FUNCTION_BLOCK "FB5002_SafetyDoorV1"   // FB5002, SCL
{ S7_Optimized_Access := 'TRUE' }
// ============================================================
//  Block: FB5002_SafetyDoorV1
//  ============================================================
//  编号：FB5002
//  原始语言：LAD（规则翻译为 SCL）
//  含义：由 LAD/FBD 网络折叠生成的等效 SCL，导入前请人工复核
   VAR_INPUT
      i_DoorOverRide : Bool;   // 安全门旁路输入请求信号
      i_AutoRunning : Bool;   // 自动运行中
      i_OpenDoorPmt : Bool := TRUE;   // 开门/旁路条件
      EMMode : Bool;   // 紧急停止模式
   END_VAR
   VAR_OUTPUT
      o_DoorOverRideRelayOn : Bool;   // 安全门旁路继电器输出
      o_DoorLockRelayON : Bool;   // 安全门线圈锁定继电器输出
      o_DoorOverRideLight : Bool;   // 安全门旁路指示灯
      o_PromptDoorOverRideStartIng : Bool;   // 开始安全门旁路,等待各流程结束!
      o_PromptDoorOveRideStarted : Bool;   // 安全门旁路，注意安全！
      o_PromptDoorLockFail : Bool;   // 安全门电磁线圈锁定失败！
   END_VAR
   VAR
      TP_DoorInsert : Array[1..8] of Bool;   // 静态变量
      TP_DoorUnLock : Array[1..8] of Bool;   // 静态变量
      AtDoorUnLock : Byte;   // 静态变量
      Aux : Struct   // 静态变量
         DT1 : Bool;   // 静态变量
         DT2 : Bool;   // 静态变量
         DT3 : Bool;   // 静态变量
         DT4 : Bool;   // 静态变量
         PromptPls : Bool;   // 静态变量
         sp : Int;   // 静态变量
      END_STRUCT;
      LastAddr : Int := 8;   // 静态变量
   END_VAR
BEGIN

   // ---------- 网络 1 ----------
   // 标题：旁路提示
   // 含义：条件 ((#i_DoorOverRide AND NOT (#EMMode)) AND NOT (#i_AutoRunning)) AND #i_OpenDoorPmt 成立时，将 TRUE 传送到 #o_DoorOverRideRelayOn
   IF ((#i_DoorOverRide AND NOT (#EMMode)) AND NOT (#i_AutoRunning)) AND #i_OpenDoorPmt THEN
       #o_DoorOverRideRelayOn := TRUE;
   END_IF;
   // 含义：条件 (((#i_DoorOverRide AND NOT (#EMMode)) AND NOT (#i_AutoRunning)) AND #i_OpenDoorPmt) AND #Aux.DT2 成立时，将 FALSE 传送到 #o_DoorLockRelayON
   IF (((#i_DoorOverRide AND NOT (#EMMode)) AND NOT (#i_AutoRunning)) AND #i_OpenDoorPmt) AND #Aux.DT2 THEN
       #o_DoorLockRelayON := FALSE;
   END_IF;
   // 含义：将 (((((#i_DoorOverRide AND NOT (#EMMode)) AND NOT (#i_AutoRunning)) AND #i_OpenDoorPmt) AND "DB1000_StdSignal".PLS.PS10) OR ((((#i_DoorOverRide AND NOT (#EMMode)) AND NOT (#i_AutoRunning)) AND #i_OpenDoorPmt) AND #Aux.DT2)) AND #Aux.DT1 赋给 #Aux.DT2
   #Aux.DT2 := (((((#i_DoorOverRide AND NOT (#EMMode)) AND NOT (#i_AutoRunning)) AND #i_OpenDoorPmt) AND "DB1000_StdSignal".PLS.PS10) OR ((((#i_DoorOverRide AND NOT (#EMMode)) AND NOT (#i_AutoRunning)) AND #i_OpenDoorPmt) AND #Aux.DT2)) AND #Aux.DT1;
   // 含义：将 ((((#i_DoorOverRide AND NOT (#EMMode)) AND NOT (#i_AutoRunning)) AND #i_OpenDoorPmt) AND "DB1000_StdSignal".PLS.PS10) OR ((((#i_DoorOverRide AND NOT (#EMMode)) AND NOT (#i_AutoRunning)) AND #i_OpenDoorPmt) AND #Aux.DT1) 赋给 #Aux.DT1
   #Aux.DT1 := ((((#i_DoorOverRide AND NOT (#EMMode)) AND NOT (#i_AutoRunning)) AND #i_OpenDoorPmt) AND "DB1000_StdSignal".PLS.PS10) OR ((((#i_DoorOverRide AND NOT (#EMMode)) AND NOT (#i_AutoRunning)) AND #i_OpenDoorPmt) AND #Aux.DT1);

   // ---------- 网络 2 ----------
   // 标题：旁路关闭
   // 含义：条件 ((NOT (#i_DoorOverRide) AND (#AtDoorUnLock = 16#00))) AND #Aux.DT4 成立时，将 FALSE 传送到 #o_DoorOverRideRelayOn
   IF ((NOT (#i_DoorOverRide) AND (#AtDoorUnLock = 16#00))) AND #Aux.DT4 THEN
       #o_DoorOverRideRelayOn := FALSE;
   END_IF;
   // 含义：将 ((((NOT (#i_DoorOverRide) AND (#AtDoorUnLock = 16#00))) AND NOT ("DB1000_StdSignal".PLS.PS10)) OR (((NOT (#i_DoorOverRide) AND (#AtDoorUnLock = 16#00))) AND #Aux.DT4)) AND #Aux.DT3 赋给 #Aux.DT4
   #Aux.DT4 := ((((NOT (#i_DoorOverRide) AND (#AtDoorUnLock = 16#00))) AND NOT ("DB1000_StdSignal".PLS.PS10)) OR (((NOT (#i_DoorOverRide) AND (#AtDoorUnLock = 16#00))) AND #Aux.DT4)) AND #Aux.DT3;
   // 含义：将 (((NOT (#i_DoorOverRide) AND (#AtDoorUnLock = 16#00))) AND "DB1000_StdSignal".PLS.PS10) OR (((NOT (#i_DoorOverRide) AND (#AtDoorUnLock = 16#00))) AND #Aux.DT3) 赋给 #Aux.DT3
   #Aux.DT3 := (((NOT (#i_DoorOverRide) AND (#AtDoorUnLock = 16#00))) AND "DB1000_StdSignal".PLS.PS10) OR (((NOT (#i_DoorOverRide) AND (#AtDoorUnLock = 16#00))) AND #Aux.DT3);
   // 含义：条件 NOT (#i_DoorOverRide) 成立时，将 TRUE 传送到 #o_DoorLockRelayON
   IF NOT (#i_DoorOverRide) THEN
       #o_DoorLockRelayON := TRUE;
   END_IF;

   // ---------- 网络 3 ----------
   // 标题：安全门旁路继电器输出
   // 含义：条件 #EMMode 成立时，将 FALSE 传送到 #o_DoorOverRideRelayOn
   IF #EMMode THEN
       #o_DoorOverRideRelayOn := FALSE;
   END_IF;

   // ---------- 网络 4 ----------
   // 标题：安全门旁路指示灯
   // 含义：将 #i_DoorOverRide AND NOT (#o_DoorOverRideRelayOn) 赋给 #o_PromptDoorOverRideStartIng
   #o_PromptDoorOverRideStartIng := #i_DoorOverRide AND NOT (#o_DoorOverRideRelayOn);
   // 含义：将 #i_DoorOverRide AND #o_DoorOverRideRelayOn 赋给 #o_PromptDoorOveRideStarted
   #o_PromptDoorOveRideStarted := #i_DoorOverRide AND #o_DoorOverRideRelayOn;
   // 含义：将 ((NOT (#EMMode) AND NOT (#i_DoorOverRide)) AND (#AtDoorUnLock <> 16#00)) 赋给 #o_PromptDoorLockFail
   #o_PromptDoorLockFail := ((NOT (#EMMode) AND NOT (#i_DoorOverRide)) AND (#AtDoorUnLock <> 16#00));
   // 含义：将 (NOT (#EMMode) AND (#AtDoorUnLock <> 16#00)) 赋给 #o_DoorOverRideLight
   #o_DoorOverRideLight := (NOT (#EMMode) AND (#AtDoorUnLock <> 16#00));
   // 含义：条件 #EMMode AND #i_DoorOverRide 成立时，将 TRUE 传送到 #o_DoorOverRideLight
   IF #EMMode AND #i_DoorOverRide THEN
       #o_DoorOverRideLight := TRUE;
   END_IF;
END_FUNCTION_BLOCK

FUNCTION_BLOCK "FB5004_ProdCycleTime"   // FB5004, SCL
{ S7_Optimized_Access := 'TRUE' }
// ============================================================
//  Block: FB5004_ProdCycleTime
//  ============================================================
//  编号：FB5004
//  原始语言：LAD（规则翻译为 SCL）
//  含义：由 LAD/FBD 网络折叠生成的等效 SCL，导入前请人工复核
   VAR_INPUT
      StepStart : Bool;   // 自动循环启动
   END_VAR
   VAR
      CycleTime_Net : Time;   // 机器运行时间
      CycleTime_Total : Time;   // 本次启动到下次启动时间(运行结束时更新）
      Aux : Struct   // 静态变量
         StartPls : Bool;   // 静态变量
         EndPls : Bool;   // 静态变量
         sp : Byte;   // 静态变量
         StartTime : Time_Of_Day;   // 静态变量
         LastEndTime : Time_Of_Day;   // 静态变量
      END_STRUCT;
   END_VAR
BEGIN
END_FUNCTION_BLOCK

FUNCTION_BLOCK "FB5005_ProdCounter"   // FB5005, SCL
{ S7_Optimized_Access := 'TRUE' }
// ============================================================
//  Block: FB5005_ProdCounter
//  ============================================================
//  编号：FB5005
//  原始语言：LAD（规则翻译为 SCL）
//  含义：由 LAD/FBD 网络折叠生成的等效 SCL，导入前请人工复核
   VAR_INPUT
      i_OKPartPrompt : Bool;   // 合格标志位
      i_NGPartPrompt : Bool;   // 不合格标志位
      i_ClearCounter : Bool;   // 清零功能
      i_ClearSuccessiveNGErr : Bool;   // 清除连续3件不合格报警
      SuccessiveNGCounterLimit : Int := 3;   // 连续不合格上限
      TotalNGCounterLimit : Int := 10;   // 不合格数量上限
   END_VAR
   VAR_OUTPUT
      o_SeccessiveNGErr : Bool;   // 连续3件不合格，请复位
      o_NGCounterLimitErr : Bool;   // 输出参数
   END_VAR
   VAR
      OKPart : Int;   // 合格量总计
      NGPart : Int;   // 不合格量总计
      Total : Int;   // 所有产量总计
      Aux : Struct   // 静态变量
         OKPls : Bool;   // 静态变量
         NGPls : Bool;   // 静态变量
         NGPart : Int;   // 一段时间内xxx件不合格
         SuccessiveNGCounter : Int;   // 静态变量
      END_STRUCT;
   END_VAR
BEGIN
END_FUNCTION_BLOCK

// folder: 001_KL_Standard_FB/098_KL_Lib

FUNCTION "FC_BlockMove" : Void   // FC1204, SCL
{ S7_Optimized_Access := 'FALSE' }
AUTHOR : czm
FAMILY : 通用
VERSION : 0.1
   VAR_INPUT
      srcDBNo : DB_ANY;   // 源数据的DB号
      srcType : Char;   // 源数据类型,默认是DB
      srcOffset : DInt;   // 源数据的偏移量(byte)
      dstDBNo : DB_ANY;   // 目标数据的DB号
      dstOffset : DInt;   // 目标数据的偏移量
      move_len : Int;   // 待移动的字节数目
   END_VAR
   VAR_TEMP
      area_src1 : Byte;
      area_dest1 : Byte;
   END_VAR
BEGIN
   IF #srcType = 'I' OR #srcType = 'i' THEN  //判断源目标的输入类型；
     #area_src1 := 16#81;
   ELSIF #srcType = 'Q' OR #srcType = 'q' THEN
     #area_src1 := 16#82;
   ELSIF #srcType = 'M' OR #srcType = 'm' THEN
     #area_src1 := 16#83;  
   ELSE
     #area_src1 := 16#84;
   END_IF;  //判断源目标的输入类型；



   POKE_BLK(area_src:= #area_src1,
            dbNumber_src:=#srcDBNo,
            byteOffset_src:=#srcOffset,
            area_dest:=16#84,
            dbNumber_dest:=#dstDBNo,
            byteOffset_dest:=#dstOffset,
            count:=#move_len
            );
END_FUNCTION

// folder: 002_Err_Prompt_Handle

FUNCTION_BLOCK "FB1140_Message"   // FB1140, SCL
{ S7_Optimized_Access := 'TRUE' }
// ============================================================
//  Block: FB1140_Message
//  ============================================================
//  编号：FB1140
//  原始语言：LAD（规则翻译为 SCL）
//  含义：由 LAD/FBD 网络折叠生成的等效 SCL，导入前请人工复核
   VAR_INPUT
      i_MaxSubStationNO : Int;   // 输入参数
      AllMode : Bool;   // 输入参数
   END_VAR
   VAR_OUTPUT
      o_Err : Bool;   // DB_Err任意一位=On
      o_NotPmtToStart : Bool;   // DB_PromptStartNotPmt任意一位=On
      o_SubErrorPresent : Struct   // 各子工位存在故障，用于识别各个子站是否需要回原点
         Public : Bool;   // 输出参数
         ST01 : Bool;   // 输出参数
         ST02 : Bool;   // 输出参数
         ST03 : Bool;   // 输出参数
         ST04 : Bool;   // 输出参数
         ST05 : Bool;   // 输出参数
         ST06 : Bool;   // 输出参数
         ST07 : Bool;   // 输出参数
         ST08 : Bool;   // 输出参数
         ST10 : Bool;   // 输出参数
         ST11 : Bool;   // 输出参数
      END_STRUCT;
      At_O_SubErrPresent : Word;   // 输出参数
      o_SubNotPmtToStart : Struct   // 输出参数
         Public : Bool;   // 输出参数
         ST01 : Bool;   // 输出参数
         ST02 : Bool;   // 输出参数
         ST03 : Bool;   // 输出参数
         ST04 : Bool;   // 输出参数
         ST05 : Bool;   // 输出参数
         ST06 : Bool;   // 输出参数
         ST07 : Bool;   // 输出参数
         ST08 : Bool;   // 输出参数
         ST10 : Bool;   // 输出参数
         ST11 : Bool;   // 输出参数
      END_STRUCT;
      At_O_SubNotPmtToStart : Word;   // 输出参数
      PromptValue : Int;   // 总的提示信息
      o_PromptValueArray : Array[0..31] of Int;   // 各个子工位的提示信息
      o_ErrPresent : Bool;   // 输出参数
      o_NotPmtToStartPresent : Bool;   // 输出参数
      o_ErrorPresentArray : Array[0..31] of Bool;   // 输出参数
      o_NotPmtToStartPresentArray : Array[0..31] of Bool;   // 输出参数
   END_VAR
   VAR
      xFB : "FB1141_Prompt";   // 静态变量
      Para : Struct   // 静态变量
         StartDBNO : Int;   // 静态变量
         DBLoopCounter : Int;   // 静态变量
         DBMessage_Gap : Int;   // 静态变量
      END_STRUCT;
      Para_ReserveLength : Struct   // 静态变量
         DB_PromptFree : Array[0..31] of Int;   // 静态变量
         DB_PromptStartNotPmt : Array[0..31] of Int;   // 静态变量
         DB_PromptErr : Array[0..31] of Int;   // 静态变量
      END_STRUCT;
      xAux : Struct   // 静态变量
         AnyBitOnPresentArray : Array[0..2, 0..31] of Bool;   // 静态变量
         AnyBitOnPresent : Array[0..2] of Bool;   // 静态变量
         o_PromptValueArray : Array[0..2, 0..31] of Int;   // 静态变量
         BakeArray : Array[0..2, 0..31] of Struct   // 静态变量
            ScanFinished : Bool;   // 静态变量
            PromptValueBake : Int;   // 静态变量
         END_STRUCT;
         DB_StationShift : Array[0..2] of Int;   // 静态变量
         ParaSubStationStartByteNO : Array[0..2, 0..31] of Int;   // 静态变量
         o_W_ErrPresentArray : DWord;   // 静态变量
         o_W_NotPmtToStartPresentArray : DWord;   // 静态变量
         DBNO : Int;   // 静态变量
         SubStep : Int;   // 静态变量
         JumpStepNO : Int;   // 静态变量
         SubStation : Int;   // 静态变量
         DBNumber : Int;   // 静态变量
      END_STRUCT;
      sp : Array[0..113] of Byte;   // 静态变量
      LastAddr : Int;   // 静态变量
   END_VAR
BEGIN

   // ---------- 网络 1 ----------
   // 含义：调用定时器实例 #xFB
   #xFB(i_MaxSubStationNO := 2,
        o_ErrPresent => #o_Err,
        o_NotPmtToStartPresent => #o_NotPmtToStart,
        PromptValue => #PromptValue,
        o_PromptValueArray => #o_PromptValueArray);

   // ---------- 网络 2 ----------
   // 标题：Word to Struct；
   // 含义：将 #xFB.xAux.o_W_ErrPresentArray 赋给 #At_O_SubErrPresent
   #At_O_SubErrPresent := #xFB.xAux.o_W_ErrPresentArray;
   // 含义：将 #xFB.xAux.o_W_NotPmtToStartPresentArray 赋给 #At_O_SubNotPmtToStart
   #At_O_SubNotPmtToStart := #xFB.xAux.o_W_NotPmtToStartPresentArray;
   // 含义：将 #PromptValue 赋给 "DB1900_Communication_PC".Send.PromptValue
   "DB1900_Communication_PC".Send.PromptValue := #PromptValue;

   // ---------- 网络 3 ----------
   // （空白网络）
END_FUNCTION_BLOCK

FUNCTION_BLOCK "FB1142_TypeChangePrompt"   // FB1142, SCL
{ S7_Optimized_Access := 'TRUE' }
// ============================================================
//  Block: FB1142_TypeChangePrompt
//  ============================================================
//  编号：FB1142
//  原始语言：LAD（规则翻译为 SCL）
//  含义：注释：跳出自动程序，除了强制停止外，断电重启
   VAR_INPUT
      ManMode : Bool;   // 手动模式
      Pulse_En : Bool;   // 输入参数
      PromptSourceDW : DWord;   // 输入参数
   END_VAR
   VAR_OUTPUT
      PromptValue : Int;   // 输出参数
   END_VAR
   VAR
      TP_Cmd : Word;   // 静态变量
      CmdAuto : Struct   // 静态变量
         StartTP : Bool;   // 开始换型按钮
         EndTP : Bool;   // 终止换型按钮
         OKTp : Bool;   // 确认按钮
         CancelTP : Bool;   // 取消按钮
      END_STRUCT;
      AtCmdAuto : Word;   // 静态变量
      CmdMid : Struct   // 静态变量
         StartTP : Bool;   // 开始换型按钮
         EndTP : Bool;   // 终止换型按钮
         OKTp : Bool;   // 确认按钮
         CancelTP : Bool;   // 取消按钮
      END_STRUCT;
      AtCmdMid : Word;   // 静态变量
      Status : Struct   // 静态变量
         PromptValue : Int;   // 静态变量
      END_STRUCT;
      TypeChangeStep : Struct   // 静态变量
         Start : Bool;   // 静态变量
         End : Bool;   // 静态变量
         ErrEnd : Bool;   // 静态变量
         Step1 : Bool;   // 静态变量
         Step2 : Bool;   // 静态变量
         Step3 : Bool;   // 静态变量
         Step4 : Bool;   // 静态变量
         Step5 : Bool;   // 静态变量
         Step6 : Bool;   // 静态变量
         Step7 : Bool;   // 静态变量
         Step8 : Bool;   // 静态变量
         Step9 : Bool;   // 静态变量
         Step10 : Bool;   // 静态变量
         Step11 : Bool;   // 静态变量
         Step12 : Bool;   // 静态变量
         Step13 : Bool;   // 静态变量
         Step14 : Bool;   // 静态变量
         Step15 : Bool;   // 静态变量
         Step16 : Bool;   // 静态变量
         Step17 : Bool;   // 静态变量
         Step18 : Bool;   // 静态变量
         Step19 : Bool;   // 静态变量
         Step20 : Bool;   // 静态变量
         Step21 : Bool;   // 静态变量
         Step22 : Bool;   // 静态变量
         Step23 : Bool;   // 静态变量
         Step24 : Bool;   // 静态变量
         Step25 : Bool;   // 静态变量
         Step26 : Bool;   // 静态变量
         Step27 : Bool;   // 静态变量
         Step28 : Bool;   // 静态变量
         Step29 : Bool;   // 静态变量
         Step30 : Bool;   // 静态变量
         Step31 : Bool;   // 静态变量
         Step32 : Bool;   // 静态变量
         Step33 : Bool;   // 静态变量
         Step34 : Bool;   // 静态变量
         Step35 : Bool;   // 静态变量
         Step36 : Bool;   // 静态变量
         Step37 : Bool;   // 静态变量
         JumpS1 : Bool;   // 静态变量
         JumpS2 : Bool;   // 静态变量
         JumpS3 : Bool;   // 静态变量
         JumpS4 : Bool;   // 静态变量
      END_STRUCT;
      Aux : Struct   // 静态变量
         TypeName : String[20];   // 静态变量
      END_STRUCT;
      InfoStruct : Struct   // 静态变量
         ComfirmTypeChange : Bool;   // 确认是否开始换型.....
         ManMode : Bool;   // 设备需在手动下换型.....
         HomPos : Bool;   // 设备不在原点状态，需复位回原点....
         MESSelect : Bool;   // 设备的联机模式，按确认....
         TypeSelect : Bool;   // 点击确认按钮进入型号选择画面.......
         WaitIngEnd : Bool;   // 等待Load参数结束.....
         OpenSafetyDoor : Bool;   // 请确认打开安全门......
         CloseSafetyDoor : Bool;   // 关闭安全门后，按确认....
         TypeChangeEnd : Bool;   // 点击确认，换型结束
         WaitIngScreenjump : Bool;   // 换型结束，等待页面跳转...
         SP1 : Bool;   // Info.XX
         SP2 : Bool;   // Info.XX
         SP3 : Bool;   // Info.XX
         SP4 : Bool;   // Info.XX
         SP5 : Bool;   // Info.XX
         SP6 : Bool;   // Info.XX
         SP7 : Bool;   // Info.XX
         SP8 : Bool;   // Info.XX
         SP9 : Bool;   // Info.XX
         SP10 : Bool;   // Info.XX
         SP11 : Bool;   // Info.XX
         SP12 : Bool;   // Info.XX
         SP13 : Bool;   // Info.XX
         SP14 : Bool;   // Info.XX
         SP15 : Bool;   // Info.XX
         SP16 : Bool;   // Info.XX
         SP17 : Bool;   // Info.XX
         SP18 : Bool;   // Info.XX
         SP19 : Bool;   // Info.XX
         SP20 : Bool;   // Info.XX
         SP21 : Bool;   // Info.XX
         SP22 : Bool;   // Info.XX
      END_STRUCT;
      AtInfoStruct : DWord;   // 静态变量
      FB_InfoPrompt : "FB1021_Prompt_Object";   // 静态变量
      CycleTime : Int;   // 静态变量
      PromptValueBake : Int;   // 静态变量
      ShiftBake : Int;   // 静态变量
   END_VAR
   VAR_TEMP
      T_DWORD : DWord;   // 临时变量
   END_VAR
BEGIN

   // ---------- 网络 1 ----------
   // 标题：按钮来自触摸屏，本网络无需修改
   // Word OR resolved
   // 含义：将 0 赋给 #TP_Cmd
   #TP_Cmd := 0;

   // ---------- 网络 2 ----------
   // 标题：强制结束换型，页面跳转到主画面
   // 含义：条件 #CmdMid.EndTP 成立时，将 200 传送到 "DB1001_SysMode".SubSysMode.TPSetPageNo
   IF #CmdMid.EndTP THEN
       "DB1001_SysMode".SubSysMode.TPSetPageNo := 200;
   END_IF;

   // ---------- 网络 3 ----------
   // 标题：****************Start******************************************
   // 注释：注释：跳出自动程序，除了强制停止外，断电重启
   // 含义：将 (((#CmdMid.StartTP OR #TypeChangeStep.Start) AND NOT (#CmdMid.EndTP)) AND NOT ("DB1000_StdSignal".PLS.InitialPls)) AND NOT (#TypeChangeStep.End) 赋给 #TypeChangeStep.Start
   #TypeChangeStep.Start := (((#CmdMid.StartTP OR #TypeChangeStep.Start) AND NOT (#CmdMid.EndTP)) AND NOT ("DB1000_StdSignal".PLS.InitialPls)) AND NOT (#TypeChangeStep.End);
   // 含义：条件 NOT ((((#CmdMid.StartTP OR #TypeChangeStep.Start) AND NOT (#CmdMid.EndTP)) AND NOT ("DB1000_StdSignal".PLS.InitialPls)) AND NOT (#TypeChangeStep.End)) 成立时，将 FALSE 传送到 #TypeChangeStep.ErrEnd
   IF NOT ((((#CmdMid.StartTP OR #TypeChangeStep.Start) AND NOT (#CmdMid.EndTP)) AND NOT ("DB1000_StdSignal".PLS.InitialPls)) AND NOT (#TypeChangeStep.End)) THEN
       #TypeChangeStep.ErrEnd := FALSE;
   END_IF;
   // 含义：条件 NOT ((((#CmdMid.StartTP OR #TypeChangeStep.Start) AND NOT (#CmdMid.EndTP)) AND NOT ("DB1000_StdSignal".PLS.InitialPls)) AND NOT (#TypeChangeStep.End)) 成立时，将 FALSE 传送到 #InfoStruct.HomPos
   IF NOT ((((#CmdMid.StartTP OR #TypeChangeStep.Start) AND NOT (#CmdMid.EndTP)) AND NOT ("DB1000_StdSignal".PLS.InitialPls)) AND NOT (#TypeChangeStep.End)) THEN
       #InfoStruct.HomPos := FALSE;
   END_IF;
   // 含义：条件 (((#CmdMid.StartTP OR #TypeChangeStep.Start) AND NOT (#CmdMid.EndTP)) AND NOT ("DB1000_StdSignal".PLS.InitialPls)) AND NOT (#TypeChangeStep.End) 成立时，将 FALSE 传送到 #CmdMid.StartTP
   IF (((#CmdMid.StartTP OR #TypeChangeStep.Start) AND NOT (#CmdMid.EndTP)) AND NOT ("DB1000_StdSignal".PLS.InitialPls)) AND NOT (#TypeChangeStep.End) THEN
       #CmdMid.StartTP := FALSE;
   END_IF;

   // ---------- 网络 4 ----------
   // 标题：StepS1,进入换型画面
   // 注释：注释：强制进入换型界面
   // String Move resolved
   // 含义：条件 ((#TypeChangeStep.Start AND NOT (#TypeChangeStep.ErrEnd)) AND ("DB1001_SysMode".SubSysMode.TPCurPageType <> 400)) 成立时，将 400 传送到 "DB1001_SysMode".SubSysMode.TPSetPageNo
   IF ((#TypeChangeStep.Start AND NOT (#TypeChangeStep.ErrEnd)) AND ("DB1001_SysMode".SubSysMode.TPCurPageType <> 400)) THEN
       "DB1001_SysMode".SubSysMode.TPSetPageNo := 400;
   END_IF;
   // 含义：将 #TypeChangeStep.Start AND NOT (#TypeChangeStep.ErrEnd) 赋给 #TypeChangeStep.Step1
   #TypeChangeStep.Step1 := #TypeChangeStep.Start AND NOT (#TypeChangeStep.ErrEnd);

   // ---------- 网络 5 ----------
   // 标题：确定是否开始确认换型
   // 含义：将 #TypeChangeStep.Step1 AND NOT (#TypeChangeStep.Step2) 赋给 #InfoStruct.ComfirmTypeChange
   #InfoStruct.ComfirmTypeChange := #TypeChangeStep.Step1 AND NOT (#TypeChangeStep.Step2);
   // 含义：条件 (#TypeChangeStep.Step1 AND NOT (#TypeChangeStep.Step2)) AND #CmdMid.CancelTP 成立时，将 TRUE 传送到 #TypeChangeStep.ErrEnd
   IF (#TypeChangeStep.Step1 AND NOT (#TypeChangeStep.Step2)) AND #CmdMid.CancelTP THEN
       #TypeChangeStep.ErrEnd := TRUE;
   END_IF;
   // 含义：将 ((#TypeChangeStep.Step1 AND #CmdMid.OKTp) AND NOT (#TypeChangeStep.ErrEnd)) OR (#TypeChangeStep.Step1 AND #TypeChangeStep.Step2) 赋给 #TypeChangeStep.Step2
   #TypeChangeStep.Step2 := ((#TypeChangeStep.Step1 AND #CmdMid.OKTp) AND NOT (#TypeChangeStep.ErrEnd)) OR (#TypeChangeStep.Step1 AND #TypeChangeStep.Step2);

   // ---------- 网络 6 ----------
   // 标题：设备需在手动模式下换型
   // 注释：注：换型过程中，必须一直在手动情况下
   // 含义：将 #TypeChangeStep.Step2 AND NOT (#TypeChangeStep.Step3) 赋给 #InfoStruct.ManMode
   #InfoStruct.ManMode := #TypeChangeStep.Step2 AND NOT (#TypeChangeStep.Step3);
   // 含义：将 #TypeChangeStep.Step2 AND #ManMode 赋给 #TypeChangeStep.Step3
   #TypeChangeStep.Step3 := #TypeChangeStep.Step2 AND #ManMode;

   // ---------- 网络 7 ----------
   // 标题：备用步
   // 含义：当 #TypeChangeStep.Step3 为 TRUE 时置位 #TypeChangeStep.Step4，否则复位（触点→线圈）
   IF #TypeChangeStep.Step3 THEN
       #TypeChangeStep.Step4 := TRUE;
   ELSE
       #TypeChangeStep.Step4 := FALSE;
   END_IF;

   // ---------- 网络 8 ----------
   // 标题：设备提示回原点
   // 含义：当 #TypeChangeStep.Step4 为 TRUE 时置位 #TypeChangeStep.Step5，否则复位（触点→线圈）
   IF #TypeChangeStep.Step4 THEN
       #TypeChangeStep.Step5 := TRUE;
   ELSE
       #TypeChangeStep.Step5 := FALSE;
   END_IF;

   // ---------- 网络 9 ----------
   // 标题：复位提示，一些特殊的处理
   // 含义：条件 #TypeChangeStep.Step5 AND NOT (#TypeChangeStep.Step6) 成立时，将 FALSE 传送到 #InfoStruct.HomPos
   IF #TypeChangeStep.Step5 AND NOT (#TypeChangeStep.Step6) THEN
       #InfoStruct.HomPos := FALSE;
   END_IF;
   // 含义：当 #TypeChangeStep.Step5 为 TRUE 时置位 #TypeChangeStep.Step6，否则复位（触点→线圈）
   IF #TypeChangeStep.Step5 THEN
       #TypeChangeStep.Step6 := TRUE;
   ELSE
       #TypeChangeStep.Step6 := FALSE;
   END_IF;

   // ---------- 网络 10 ----------
   // 标题：确认设备的状态，单机OR联机
   // 含义：将 #TypeChangeStep.Step6 AND NOT (#TypeChangeStep.Step7) 赋给 #InfoStruct.MESSelect
   #InfoStruct.MESSelect := #TypeChangeStep.Step6 AND NOT (#TypeChangeStep.Step7);
   // 含义：将 (#TypeChangeStep.Step6 AND #CmdMid.OKTp) OR (#TypeChangeStep.Step6 AND #TypeChangeStep.Step7) 赋给 #TypeChangeStep.Step7
   #TypeChangeStep.Step7 := (#TypeChangeStep.Step6 AND #CmdMid.OKTp) OR (#TypeChangeStep.Step6 AND #TypeChangeStep.Step7);

   // ---------- 网络 11 ----------
   // 标题：即将进入换型界面,点击确认
   // 含义：将 #TypeChangeStep.Step7 AND NOT (#TypeChangeStep.Step8) 赋给 #InfoStruct.TypeSelect
   #InfoStruct.TypeSelect := #TypeChangeStep.Step7 AND NOT (#TypeChangeStep.Step8);
   // 含义：条件 (#TypeChangeStep.Step7 AND NOT (#TypeChangeStep.Step8)) AND #CmdMid.OKTp 成立时，将 401 传送到 "DB1001_SysMode".SubSysMode.TPSetPageNo
   IF (#TypeChangeStep.Step7 AND NOT (#TypeChangeStep.Step8)) AND #CmdMid.OKTp THEN
       "DB1001_SysMode".SubSysMode.TPSetPageNo := 401;
   END_IF;
   // 含义：将 (#TypeChangeStep.Step7 AND #CmdMid.OKTp) OR (#TypeChangeStep.Step7 AND #TypeChangeStep.Step8) 赋给 #TypeChangeStep.Step8
   #TypeChangeStep.Step8 := (#TypeChangeStep.Step7 AND #CmdMid.OKTp) OR (#TypeChangeStep.Step7 AND #TypeChangeStep.Step8);

   // ---------- 网络 12 ----------
   // 标题：进入换型界面"DB_Parameter".CmdMid.TypeConfirm
   // 含义：条件 ((#TypeChangeStep.Step8 AND NOT (#TypeChangeStep.Step10)) AND ("DB1001_SysMode".SubSysMode.TPSetPageNo <> 401)) 成立时，将 499 传送到 "DB1001_SysMode".SubSysMode.TPSetPageNo
   IF ((#TypeChangeStep.Step8 AND NOT (#TypeChangeStep.Step10)) AND ("DB1001_SysMode".SubSysMode.TPSetPageNo <> 401)) THEN
       "DB1001_SysMode".SubSysMode.TPSetPageNo := 499;
   END_IF;
   // 含义：将 (#TypeChangeStep.Step8 AND TRUE) OR (#TypeChangeStep.Step8 AND #TypeChangeStep.Step10) 赋给 #TypeChangeStep.Step10
   #TypeChangeStep.Step10 := (#TypeChangeStep.Step8 AND TRUE) OR (#TypeChangeStep.Step8 AND #TypeChangeStep.Step10);

   // ---------- 网络 13 ----------
   // 标题：打开安全门
   // 含义：将 #TypeChangeStep.Step10 AND NOT (#TypeChangeStep.Step11) 赋给 #InfoStruct.OpenSafetyDoor
   #InfoStruct.OpenSafetyDoor := #TypeChangeStep.Step10 AND NOT (#TypeChangeStep.Step11);
   // 含义：条件 #TypeChangeStep.Step10 AND NOT (#TypeChangeStep.Step11) 成立时，将 400 传送到 "DB1001_SysMode".SubSysMode.TPSetPageNo
   IF #TypeChangeStep.Step10 AND NOT (#TypeChangeStep.Step11) THEN
       "DB1001_SysMode".SubSysMode.TPSetPageNo := 400;
   END_IF;
   // 含义：将 (#TypeChangeStep.Step10 AND #CmdMid.OKTp) OR (#TypeChangeStep.Step10 AND #TypeChangeStep.Step11) 赋给 #TypeChangeStep.Step11
   #TypeChangeStep.Step11 := (#TypeChangeStep.Step10 AND #CmdMid.OKTp) OR (#TypeChangeStep.Step10 AND #TypeChangeStep.Step11);

   // ---------- 网络 14 ----------
   // 标题：换夹具提示信息
   // 含义：当 #TypeChangeStep.Step11 为 TRUE 时置位 #TypeChangeStep.Step12，否则复位（触点→线圈）
   IF #TypeChangeStep.Step11 THEN
       #TypeChangeStep.Step12 := TRUE;
   ELSE
       #TypeChangeStep.Step12 := FALSE;
   END_IF;

   // ---------- 网络 15 ----------
   // 标题：关闭安全门
   // 含义：将 #TypeChangeStep.Step12 AND NOT (#TypeChangeStep.Step28) 赋给 #InfoStruct.CloseSafetyDoor
   #InfoStruct.CloseSafetyDoor := #TypeChangeStep.Step12 AND NOT (#TypeChangeStep.Step28);
   // 含义：将 (#TypeChangeStep.Step12 AND #CmdMid.OKTp) OR (#TypeChangeStep.Step12 AND #TypeChangeStep.Step28) 赋给 #TypeChangeStep.Step28
   #TypeChangeStep.Step28 := (#TypeChangeStep.Step12 AND #CmdMid.OKTp) OR (#TypeChangeStep.Step12 AND #TypeChangeStep.Step28);

   // ---------- 网络 16 ----------
   // 标题：提示回原点
   // 含义：当 #TypeChangeStep.Step28 为 TRUE 时置位 #TypeChangeStep.Step30，否则复位（触点→线圈）
   IF #TypeChangeStep.Step28 THEN
       #TypeChangeStep.Step30 := TRUE;
   ELSE
       #TypeChangeStep.Step30 := FALSE;
   END_IF;

   // ---------- 网络 17 ----------
   // 标题：换型结束
   // 含义：将 (#TypeChangeStep.Step30 OR #TypeChangeStep.ErrEnd) AND NOT (#TypeChangeStep.Step32) 赋给 #InfoStruct.TypeChangeEnd
   #InfoStruct.TypeChangeEnd := (#TypeChangeStep.Step30 OR #TypeChangeStep.ErrEnd) AND NOT (#TypeChangeStep.Step32);
   // 含义：将 #TypeChangeStep.Step30 OR #TypeChangeStep.ErrEnd 赋给 #TypeChangeStep.Step32
   #TypeChangeStep.Step32 := #TypeChangeStep.Step30 OR #TypeChangeStep.ErrEnd;

   // ---------- 网络 18 ----------
   // 标题：切换到自动画面
   // 含义：条件 #TypeChangeStep.Step32 AND NOT (#TypeChangeStep.Step33) 成立时，将 200 传送到 "DB1001_SysMode".SubSysMode.TPSetPageNo
   IF #TypeChangeStep.Step32 AND NOT (#TypeChangeStep.Step33) THEN
       "DB1001_SysMode".SubSysMode.TPSetPageNo := 200;
   END_IF;
   // 含义：将 #TypeChangeStep.Step32 AND NOT (#TypeChangeStep.Step33) 赋给 #InfoStruct.WaitIngScreenjump
   #InfoStruct.WaitIngScreenjump := #TypeChangeStep.Step32 AND NOT (#TypeChangeStep.Step33);
   // 含义：当 #TypeChangeStep.Step32 为 TRUE 时置位 #TypeChangeStep.End，否则复位（触点→线圈）
   IF #TypeChangeStep.Step32 THEN
       #TypeChangeStep.End := TRUE;
   ELSE
       #TypeChangeStep.End := FALSE;
   END_IF;

   // ---------- 网络 19 ----------
   // 标题：InfoStruct --> Prompt
   // 含义：调用定时器实例 #FB_InfoPrompt
   #FB_InfoPrompt(Pulse_En := "DB1000_StdSignal".PLS.PS10,
                  PromptSourceDW := #AtInfoStruct,
                  PromptValue => #Status.PromptValue);

   // ---------- 网络 20 ----------
   // （空白网络）
END_FUNCTION_BLOCK

// folder: 003_HomeStep

FUNCTION_BLOCK "FB1040_HomePos"   // FB1040, SCL
{ S7_Optimized_Access := 'TRUE' }
// ============================================================
//  Block: FB1040_HomePos
//  ============================================================
//  编号：FB1040
//  原始语言：LAD（规则翻译为 SCL）
//  含义：由 LAD/FBD 网络折叠生成的等效 SCL，导入前请人工复核
   VAR
      Status : Struct   // 状态
         Running : Bool;   // 回原点运行中
         AllStationInHomePos : Bool;   // 设备在原点位置
         AllSubStationInHomePos : Bool;   // 所有子工位在原点位置( 安全门等除外 ）
      END_STRUCT;
      MainStep : "UDT_Step";   // 回原点流程步
      EdgeDetc : Struct   // 静态变量
         JUMP : Array[0..7] of Bool;   // 静态变量
      END_STRUCT;
      StartCmd_ManMode : Bool;   // 静态变量
      StartCmd_AutoMode : Bool;   // 静态变量
      OkToStart : Bool;   // 静态变量
      HomePos : Bool;   // 静态变量
      "Do" : Bool;   // 静态变量
      Done : Bool;   // 静态变量
      PartOn : Bool;   // 静态变量
      PartOK : Bool;   // 静态变量
      PartNG : Bool;   // 静态变量
      Start : Bool;   // 静态变量
      End : Bool;   // 静态变量
      ErrEnd : Bool;   // 静态变量
      S1 : Bool;   // 静态变量
      S2 : Bool;   // 静态变量
      S3 : Bool;   // 静态变量
      S4 : Bool;   // 静态变量
      S5 : Bool;   // 静态变量
      S6 : Bool;   // 静态变量
      S7 : Bool;   // 静态变量
      S8 : Bool;   // 静态变量
      S9 : Bool;   // 静态变量
      S10 : Bool;   // 静态变量
      S11 : Bool;   // 静态变量
      S12 : Bool;   // 静态变量
      S13 : Bool;   // 静态变量
      S14 : Bool;   // 静态变量
      S15 : Bool;   // 静态变量
      S16 : Bool;   // 静态变量
      S17 : Bool;   // 静态变量
      S18 : Bool;   // 静态变量
      S19 : Bool;   // 静态变量
      S20 : Bool;   // 静态变量
      S21 : Bool;   // 静态变量
      S22 : Bool;   // 静态变量
      S23 : Bool;   // 静态变量
      S24 : Bool;   // 静态变量
      S25 : Bool;   // 静态变量
      S26 : Bool;   // 静态变量
      S27 : Bool;   // 静态变量
      S28 : Bool;   // 静态变量
      S29 : Bool;   // 静态变量
      S30 : Bool;   // 静态变量
      S31 : Bool;   // 静态变量
      S32 : Bool;   // 静态变量
      S33 : Bool;   // 静态变量
      S34 : Bool;   // 静态变量
      S35 : Bool;   // 静态变量
      S36 : Bool;   // 静态变量
      S37 : Bool;   // 静态变量
      S38 : Bool;   // 静态变量
      S39 : Bool;   // 静态变量
      S40 : Bool;   // 静态变量
      S41 : Bool;   // 静态变量
      S42 : Bool;   // 静态变量
      S43 : Bool;   // 静态变量
      S44 : Bool;   // 静态变量
      S45 : Bool;   // 静态变量
      S46 : Bool;   // 静态变量
      S47 : Bool;   // 静态变量
      S48 : Bool;   // 静态变量
      S49 : Bool;   // 静态变量
      S50 : Bool;   // 静态变量
      S51 : Bool;   // 静态变量
      S52 : Bool;   // 静态变量
      S53 : Bool;   // 静态变量
      S54 : Bool;   // 静态变量
      S55 : Bool;   // 静态变量
      S56 : Bool;   // 静态变量
      S57 : Bool;   // 静态变量
      S58 : Bool;   // 静态变量
      S59 : Bool;   // 静态变量
      S60 : Bool;   // 静态变量
      S61 : Bool;   // 静态变量
      S62 : Bool;   // 静态变量
      S63 : Bool;   // 静态变量
      S64 : Bool;   // 静态变量
      S65 : Bool;   // 静态变量
      S66 : Bool;   // 静态变量
      S67 : Bool;   // 静态变量
   END_VAR
BEGIN

   // ---------- 网络 1 ----------
   // 标题：回原点运行中
   // 含义：当 #MainStep.Start 为 TRUE 时置位 #Status.Running，否则复位（触点→线圈）
   IF #MainStep.Start THEN
       #Status.Running := TRUE;
   ELSE
       #Status.Running := FALSE;
   END_IF;

   // ---------- 网络 2 ----------
   // 标题：设备在原点位置
   // 含义：将 (((((("DB1081_ValveCall".ST01.Z01.ExtPos AND "DB1081_ValveCall".ST01.Z05.RetPos) OR ("DB1081_ValveCall".ST01.Z01.ExtPos AND NOT ("DB1081_ValveCall".ST01.Z05.ExtPos))) AND "DB1080_Component".Robot.Status.HomePos) AND "DB1081_ValveCall".ST01.Z03.RetPos) OR (((("DB1081_ValveCall".ST01.Z01.ExtPos AND "DB1081_ValveCall".ST01.Z05.RetPos) OR ("DB1081_ValveCall".ST01.Z01.ExtPos AND NOT ("DB1081_ValveCall".ST01.Z05.ExtPos))) AND "DB1080_Component".Robot.Status.HomePos) AND NOT ("DB720_KuKa_MainCtrl".Aux.AStation_ToolAtPosT.Q))) AND "DB1081_ValveCall".ST01.Z04.RetPos) OR (((((("DB1081_ValveCall".ST01.Z01.ExtPos AND "DB1081_ValveCall".ST01.Z05.RetPos) OR ("DB1081_ValveCall".ST01.Z01.ExtPos AND NOT ("DB1081_ValveCall".ST01.Z05.ExtPos))) AND "DB1080_Component".Robot.Status.HomePos) AND "DB1081_ValveCall".ST01.Z03.RetPos) OR (((("DB1081_ValveCall".ST01.Z01.ExtPos AND "DB1081_ValveCall".ST01.Z05.RetPos) OR ("DB1081_ValveCall".ST01.Z01.ExtPos AND NOT ("DB1081_ValveCall".ST01.Z05.ExtPos))) AND "DB1080_Component".Robot.Status.HomePos) AND NOT ("DB720_KuKa_MainCtrl".Aux.AStation_ToolAtPosT.Q))) AND NOT ("DB720_KuKa_MainCtrl".Aux.BStation_ToolAtPosT.Q)) 赋给 #Status.AllSubStationInHomePos
   #Status.AllSubStationInHomePos := (((((("DB1081_ValveCall".ST01.Z01.ExtPos AND "DB1081_ValveCall".ST01.Z05.RetPos) OR ("DB1081_ValveCall".ST01.Z01.ExtPos AND NOT ("DB1081_ValveCall".ST01.Z05.ExtPos))) AND "DB1080_Component".Robot.Status.HomePos) AND "DB1081_ValveCall".ST01.Z03.RetPos) OR (((("DB1081_ValveCall".ST01.Z01.ExtPos AND "DB1081_ValveCall".ST01.Z05.RetPos) OR ("DB1081_ValveCall".ST01.Z01.ExtPos AND NOT ("DB1081_ValveCall".ST01.Z05.ExtPos))) AND "DB1080_Component".Robot.Status.HomePos) AND NOT ("DB720_KuKa_MainCtrl".Aux.AStation_ToolAtPosT.Q))) AND "DB1081_ValveCall".ST01.Z04.RetPos) OR (((((("DB1081_ValveCall".ST01.Z01.ExtPos AND "DB1081_ValveCall".ST01.Z05.RetPos) OR ("DB1081_ValveCall".ST01.Z01.ExtPos AND NOT ("DB1081_ValveCall".ST01.Z05.ExtPos))) AND "DB1080_Component".Robot.Status.HomePos) AND "DB1081_ValveCall".ST01.Z03.RetPos) OR (((("DB1081_ValveCall".ST01.Z01.ExtPos AND "DB1081_ValveCall".ST01.Z05.RetPos) OR ("DB1081_ValveCall".ST01.Z01.ExtPos AND NOT ("DB1081_ValveCall".ST01.Z05.ExtPos))) AND "DB1080_Component".Robot.Status.HomePos) AND NOT ("DB720_KuKa_MainCtrl".Aux.AStation_ToolAtPosT.Q))) AND NOT ("DB720_KuKa_MainCtrl".Aux.BStation_ToolAtPosT.Q));
   // 含义：当 #Status.AllSubStationInHomePos 为 TRUE 时置位 #Status.AllStationInHomePos，否则复位（触点→线圈）
   IF #Status.AllSubStationInHomePos THEN
       #Status.AllStationInHomePos := TRUE;
   ELSE
       #Status.AllStationInHomePos := FALSE;
   END_IF;
   // 含义：将 "ManMode_M" OR "AutoMode_M" 赋给 #EdgeDetc.JUMP[0]
   #EdgeDetc.JUMP[0] := "ManMode_M" OR "AutoMode_M";
   // 含义：条件 "ManMode_M" 成立时，将 TRUE 传送到 "DB1081_ValveCall".ST01.Z05.RetAuto
   IF "ManMode_M" THEN
       "DB1081_ValveCall".ST01.Z05.RetAuto := TRUE;
   END_IF;

   // ---------- 网络 3 ----------
   // 标题：回原点开始
   // 含义：将 (((((((("ManMode_M" AND "DB1001_SysMode".SubSysMode.Mode.HomeCmd) AND NOT ("DB1080_Component".Robot.Status.Busy)) OR (("AutoMode_M" AND "DB1148_PromptBeeper".Public.ConcreteEnd) AND NOT ("DB1080_Component".Robot.Status.HomePos)) OR #MainStep.Start) AND NOT (#EdgeDetc.JUMP[0])) AND NOT (#MainStep.End)) AND NOT (#MainStep.ErrEnd)) AND NOT ("DB1080_Component".SafetyDoor.i_DoorOverRide)) AND NOT ("DB1080_Component".SafetyDoor.i_DoorOverRide)) OR (((((((("ManMode_M" AND "DB1001_SysMode".SubSysMode.Mode.HomeCmd) AND NOT ("DB1080_Component".Robot.Status.Busy)) OR (("AutoMode_M" AND "DB1148_PromptBeeper".Public.ConcreteEnd) AND NOT ("DB1080_Component".Robot.Status.HomePos)) OR #MainStep.Start) AND NOT (#EdgeDetc.JUMP[0])) AND NOT (#MainStep.End)) AND NOT (#MainStep.ErrEnd)) AND NOT ("DB1080_Component".SafetyDoor.i_DoorOverRide)) AND "DB720_KuKa_MainCtrl".StatusIn.do_FixStationToHome) OR ((((((((((("ManMode_M" AND "DB1001_SysMode".SubSysMode.Mode.HomeCmd) AND NOT ("DB1080_Component".Robot.Status.Busy)) OR (("AutoMode_M" AND "DB1148_PromptBeeper".Public.ConcreteEnd) AND NOT ("DB1080_Component".Robot.Status.HomePos)) OR #MainStep.Start) AND NOT (#EdgeDetc.JUMP[0])) AND NOT (#MainStep.End)) AND NOT (#MainStep.ErrEnd)) AND NOT ("DB1080_Component".SafetyDoor.i_DoorOverRide)) AND "BStation_ToolOn2") AND "AStation_ToolOn2") AND NOT (#Status.AllStationInHomePos)) AND "DB1081_ValveCall".ST01.Z07.ExtPos) OR (((((((((((("ManMode_M" AND "DB1001_SysMode".SubSysMode.Mode.HomeCmd) AND NOT ("DB1080_Component".Robot.Status.Busy)) OR (("AutoMode_M" AND "DB1148_PromptBeeper".Public.ConcreteEnd) AND NOT ("DB1080_Component".Robot.Status.HomePos)) OR #MainStep.Start) AND NOT (#EdgeDetc.JUMP[0])) AND NOT (#MainStep.End)) AND NOT (#MainStep.ErrEnd)) AND NOT ("DB1080_Component".SafetyDoor.i_DoorOverRide)) AND "DB1900_Communication_PC".Para.ProduceMode3) AND "IZ02RetPos") OR (((((((("ManMode_M" AND "DB1001_SysMode".SubSysMode.Mode.HomeCmd) AND NOT ("DB1080_Component".Robot.Status.Busy)) OR (("AutoMode_M" AND "DB1148_PromptBeeper".Public.ConcreteEnd) AND NOT ("DB1080_Component".Robot.Status.HomePos)) OR #MainStep.Start) AND NOT (#EdgeDetc.JUMP[0])) AND NOT (#MainStep.End)) AND NOT (#MainStep.ErrEnd)) AND NOT ("DB1080_Component".SafetyDoor.i_DoorOverRide)) AND NOT ("DB1900_Communication_PC".Para.ProduceMode3))) AND NOT (#Status.AllStationInHomePos)) AND NOT ("DB720_KuKa_MainCtrl".StatusIn.do_FixStationToHome)) 赋给 #MainStep.Start
   #MainStep.Start := (((((((("ManMode_M" AND "DB1001_SysMode".SubSysMode.Mode.HomeCmd) AND NOT ("DB1080_Component".Robot.Status.Busy)) OR (("AutoMode_M" AND "DB1148_PromptBeeper".Public.ConcreteEnd) AND NOT ("DB1080_Component".Robot.Status.HomePos)) OR #MainStep.Start) AND NOT (#EdgeDetc.JUMP[0])) AND NOT (#MainStep.End)) AND NOT (#MainStep.ErrEnd)) AND NOT ("DB1080_Component".SafetyDoor.i_DoorOverRide)) AND NOT ("DB1080_Component".SafetyDoor.i_DoorOverRide)) OR (((((((("ManMode_M" AND "DB1001_SysMode".SubSysMode.Mode.HomeCmd) AND NOT ("DB1080_Component".Robot.Status.Busy)) OR (("AutoMode_M" AND "DB1148_PromptBeeper".Public.ConcreteEnd) AND NOT ("DB1080_Component".Robot.Status.HomePos)) OR #MainStep.Start) AND NOT (#EdgeDetc.JUMP[0])) AND NOT (#MainStep.End)) AND NOT (#MainStep.ErrEnd)) AND NOT ("DB1080_Component".SafetyDoor.i_DoorOverRide)) AND "DB720_KuKa_MainCtrl".StatusIn.do_FixStationToHome) OR ((((((((((("ManMode_M" AND "DB1001_SysMode".SubSysMode.Mode.HomeCmd) AND NOT ("DB1080_Component".Robot.Status.Busy)) OR (("AutoMode_M" AND "DB1148_PromptBeeper".Public.ConcreteEnd) AND NOT ("DB1080_Component".Robot.Status.HomePos)) OR #MainStep.Start) AND NOT (#EdgeDetc.JUMP[0])) AND NOT (#MainStep.End)) AND NOT (#MainStep.ErrEnd)) AND NOT ("DB1080_Component".SafetyDoor.i_DoorOverRide)) AND "BStation_ToolOn2") AND "AStation_ToolOn2") AND NOT (#Status.AllStationInHomePos)) AND "DB1081_ValveCall".ST01.Z07.ExtPos) OR (((((((((((("ManMode_M" AND "DB1001_SysMode".SubSysMode.Mode.HomeCmd) AND NOT ("DB1080_Component".Robot.Status.Busy)) OR (("AutoMode_M" AND "DB1148_PromptBeeper".Public.ConcreteEnd) AND NOT ("DB1080_Component".Robot.Status.HomePos)) OR #MainStep.Start) AND NOT (#EdgeDetc.JUMP[0])) AND NOT (#MainStep.End)) AND NOT (#MainStep.ErrEnd)) AND NOT ("DB1080_Component".SafetyDoor.i_DoorOverRide)) AND "DB1900_Communication_PC".Para.ProduceMode3) AND "IZ02RetPos") OR (((((((("ManMode_M" AND "DB1001_SysMode".SubSysMode.Mode.HomeCmd) AND NOT ("DB1080_Component".Robot.Status.Busy)) OR (("AutoMode_M" AND "DB1148_PromptBeeper".Public.ConcreteEnd) AND NOT ("DB1080_Component".Robot.Status.HomePos)) OR #MainStep.Start) AND NOT (#EdgeDetc.JUMP[0])) AND NOT (#MainStep.End)) AND NOT (#MainStep.ErrEnd)) AND NOT ("DB1080_Component".SafetyDoor.i_DoorOverRide)) AND NOT ("DB1900_Communication_PC".Para.ProduceMode3))) AND NOT (#Status.AllStationInHomePos)) AND NOT ("DB720_KuKa_MainCtrl".StatusIn.do_FixStationToHome));

   // ---------- 网络 4 ----------
   // 标题：机器人回原点之后关枪 and Reset Robot Return Home Cmd
   // 含义：条件 ((("ManMode_M" AND "DB1080_Component".Robot.Status.HomePos) AND "DB1081_ValveCall".ST01.Z03.RetPos) AND "DB1081_ValveCall".ST01.Z04.ExtPos) OR ((("ManMode_M" AND "DB1080_Component".Robot.Status.HomePos) AND "DB1081_ValveCall".ST01.Z03.ExtPos) AND "DB1081_ValveCall".ST01.Z04.RetPos) 成立时，将 FALSE 传送到 "DB2500 Visual Chiseling".RobotRetHomeCmd_AllMode
   IF ((("ManMode_M" AND "DB1080_Component".Robot.Status.HomePos) AND "DB1081_ValveCall".ST01.Z03.RetPos) AND "DB1081_ValveCall".ST01.Z04.ExtPos) OR ((("ManMode_M" AND "DB1080_Component".Robot.Status.HomePos) AND "DB1081_ValveCall".ST01.Z03.ExtPos) AND "DB1081_ValveCall".ST01.Z04.RetPos) THEN
       "DB2500 Visual Chiseling".RobotRetHomeCmd_AllMode := FALSE;
   END_IF;
   // 含义：条件 ((("ManMode_M" AND "DB1080_Component".Robot.Status.HomePos) AND "DB1081_ValveCall".ST01.Z03.RetPos) AND "DB1081_ValveCall".ST01.Z04.ExtPos) OR ((("ManMode_M" AND "DB1080_Component".Robot.Status.HomePos) AND "DB1081_ValveCall".ST01.Z03.ExtPos) AND "DB1081_ValveCall".ST01.Z04.RetPos) OR ((("ManMode_M" AND "DB1080_Component".Robot.Status.HomePos) AND "DB1081_ValveCall".ST01.Z03.RetPos) AND "DB1081_ValveCall".ST01.Z04.RetPos) 成立时，将 FALSE 传送到 "DB2500 Visual Chiseling".RobotRetHomeCmd_AllMode
   IF ((("ManMode_M" AND "DB1080_Component".Robot.Status.HomePos) AND "DB1081_ValveCall".ST01.Z03.RetPos) AND "DB1081_ValveCall".ST01.Z04.ExtPos) OR ((("ManMode_M" AND "DB1080_Component".Robot.Status.HomePos) AND "DB1081_ValveCall".ST01.Z03.ExtPos) AND "DB1081_ValveCall".ST01.Z04.RetPos) OR ((("ManMode_M" AND "DB1080_Component".Robot.Status.HomePos) AND "DB1081_ValveCall".ST01.Z03.RetPos) AND "DB1081_ValveCall".ST01.Z04.RetPos) THEN
       "DB2500 Visual Chiseling".RobotRetHomeCmd_AllMode := FALSE;
   END_IF;

   // ---------- 网络 5 ----------
   // 标题：流程开始
   // 含义：当 #MainStep.Start 为 TRUE 时置位 #MainStep.S1，否则复位（触点→线圈）
   IF #MainStep.Start THEN
       #MainStep.S1 := TRUE;
   ELSE
       #MainStep.S1 := FALSE;
   END_IF;
   // 含义：条件 NOT (#MainStep.Start) 成立时，将 FALSE 传送到 #MainStep.ErrEnd
   IF NOT (#MainStep.Start) THEN
       #MainStep.ErrEnd := FALSE;
   END_IF;
   // 含义：条件 NOT (#MainStep.Start) 成立时，将 FALSE 传送到 #EdgeDetc.JUMP[0]
   IF NOT (#MainStep.Start) THEN
       #EdgeDetc.JUMP[0] := FALSE;
   END_IF;
   // 含义：条件 NOT (#MainStep.Start) 成立时，将 FALSE 传送到 "DB1148_PromptBeeper".Public.RetHome_Z02RetTimeOut
   IF NOT (#MainStep.Start) THEN
       "DB1148_PromptBeeper".Public.RetHome_Z02RetTimeOut := FALSE;
   END_IF;
   // 含义：条件 NOT (#MainStep.Start) 成立时，将 FALSE 传送到 "DB1148_PromptBeeper".Public.RetHome_PowerOff
   IF NOT (#MainStep.Start) THEN
       "DB1148_PromptBeeper".Public.RetHome_PowerOff := FALSE;
   END_IF;

   // ---------- 网络 6 ----------
   // 标题：推力气缸
   // 含义：条件 #MainStep.S1 AND NOT (#MainStep.S2) 成立时，将 TRUE 传送到 "DB1081_ValveCall".ST01.Z05.RetAuto
   IF #MainStep.S1 AND NOT (#MainStep.S2) THEN
       "DB1081_ValveCall".ST01.Z05.RetAuto := TRUE;
   END_IF;
   // 含义：条件 #MainStep.S1 AND NOT (#MainStep.S2) 成立时，将 TRUE 传送到 "DB1081_ValveCall".ST01.Z08.RetAuto
   IF #MainStep.S1 AND NOT (#MainStep.S2) THEN
       "DB1081_ValveCall".ST01.Z08.RetAuto := TRUE;
   END_IF;
   // 含义：将 ((#MainStep.S1 AND "DB1081_ValveCall".ST01.Z05.RetPos) AND NOT ("DB1080_Component".Robot.Status.Busy)) OR (#MainStep.S1 AND #MainStep.S2) 赋给 #MainStep.S2
   #MainStep.S2 := ((#MainStep.S1 AND "DB1081_ValveCall".ST01.Z05.RetPos) AND NOT ("DB1080_Component".Robot.Status.Busy)) OR (#MainStep.S1 AND #MainStep.S2);
   // 含义：条件 #MainStep.S1 AND "DB1042_Timer".FixtureStuckTimeOut.Q 成立时，将 TRUE 传送到 #MainStep.ErrEnd
   IF #MainStep.S1 AND "DB1042_Timer".FixtureStuckTimeOut.Q THEN
       #MainStep.ErrEnd := TRUE;
   END_IF;
   // 含义：条件 #MainStep.S1 AND "DB1042_Timer".FixtureStuckTimeOut.Q 成立时，将 TRUE 传送到 "DB1080_Component".Robot.Cmd.Auto.Stop
   IF #MainStep.S1 AND "DB1042_Timer".FixtureStuckTimeOut.Q THEN
       "DB1080_Component".Robot.Cmd.Auto.Stop := TRUE;
   END_IF;
   // 含义：条件 #MainStep.S1 AND "DB1042_Timer".FixtureStuckTimeOut.Q 成立时，将 TRUE 传送到 "DB1148_PromptBeeper".Public.BitStuckErr_Fixture
   IF #MainStep.S1 AND "DB1042_Timer".FixtureStuckTimeOut.Q THEN
       "DB1148_PromptBeeper".Public.BitStuckErr_Fixture := TRUE;
   END_IF;

   // ---------- 网络 7 ----------
   // 含义：条件 (#MainStep.S2 AND NOT (#MainStep.S6)) AND NOT ("DB1042_Timer".DrillMemory) 成立时，将 TRUE 传送到 "DB1080_Component".Robot.Cmd.Auto.GoHome
   IF (#MainStep.S2 AND NOT (#MainStep.S6)) AND NOT ("DB1042_Timer".DrillMemory) THEN
       "DB1080_Component".Robot.Cmd.Auto.GoHome := TRUE;
   END_IF;
   // 含义：条件 (#MainStep.S2 AND NOT (#MainStep.S6)) AND NOT ("DB1042_Timer".DrillMemory) 成立时，将 255 传送到 "DB1080_Component".Robot.CTRL_IN.ProgNo
   IF (#MainStep.S2 AND NOT (#MainStep.S6)) AND NOT ("DB1042_Timer".DrillMemory) THEN
       "DB1080_Component".Robot.CTRL_IN.ProgNo := 255;
   END_IF;
   // 含义：条件 (#MainStep.S2 AND NOT (#MainStep.S6)) AND "DB1042_Timer".DrillMemory 成立时，将 TRUE 传送到 "DB1081_ValveCall".ST01.Z05.ExtAuto
   IF (#MainStep.S2 AND NOT (#MainStep.S6)) AND "DB1042_Timer".DrillMemory THEN
       "DB1081_ValveCall".ST01.Z05.ExtAuto := TRUE;
   END_IF;
   // 含义：调用定时器实例 "DB1042_Timer".PowerOn_RetHome.TON
   "DB1042_Timer".PowerOn_RetHome.TON(IN := ((#MainStep.S2 AND NOT (#MainStep.S6)) AND "DB1042_Timer".DrillMemory) AND "DB1900_Communication_PC".Send.ToolPowerOn,
                                      PT := T#5S);
   // 含义：调用计数器实例 "DB1042_Timer".RetHomeHighCurrentOut.TON（上升沿计数，当前值写入 CV）
   "DB1042_Timer".RetHomeHighCurrentOut.TON(IN := ((((#MainStep.S2 AND NOT (#MainStep.S6)) AND "DB1042_Timer".DrillMemory) AND "DB1042_Timer".PowerOn_RetHome.Q) AND ("DB1900_Communication_PC".Recv.Current_2 > "DB1900_Communication_PC".Para.CurrentMaxLimit)),
                                            PT := T#100mS);
   // 含义：条件 (((#MainStep.S2 AND NOT (#MainStep.S6)) AND "DB1042_Timer".DrillMemory) AND "DB1042_Timer".PowerOn_RetHome.Q) AND NOT ("DB1042_Timer".RetHomeHighCurrentOut.Q) 成立时，将 TRUE 传送到 "DB1081_ValveCall".ST01.Z01.RetAuto
   IF (((#MainStep.S2 AND NOT (#MainStep.S6)) AND "DB1042_Timer".DrillMemory) AND "DB1042_Timer".PowerOn_RetHome.Q) AND NOT ("DB1042_Timer".RetHomeHighCurrentOut.Q) THEN
       "DB1081_ValveCall".ST01.Z01.RetAuto := TRUE;
   END_IF;
   // 含义：条件 ((((#MainStep.S2 AND NOT (#MainStep.S6)) AND "DB1042_Timer".DrillMemory) AND "DB1042_Timer".PowerOn_RetHome.Q) AND NOT ("DB1042_Timer".RetHomeHighCurrentOut.Q)) AND "DB1900_Communication_PC".Para.DrillDirection3 成立时，将 TRUE 传送到 "DB1081_ValveCall".ST01.Z02.RetAuto
   IF ((((#MainStep.S2 AND NOT (#MainStep.S6)) AND "DB1042_Timer".DrillMemory) AND "DB1042_Timer".PowerOn_RetHome.Q) AND NOT ("DB1042_Timer".RetHomeHighCurrentOut.Q)) AND "DB1900_Communication_PC".Para.DrillDirection3 THEN
       "DB1081_ValveCall".ST01.Z02.RetAuto := TRUE;
   END_IF;
   // 含义：调用定时器实例 "DB1042_Timer".RetHome_Z02TimeOut.TON
   "DB1042_Timer".RetHome_Z02TimeOut.TON(IN := ((((#MainStep.S2 AND NOT (#MainStep.S6)) AND "DB1042_Timer".DrillMemory) AND "DB1042_Timer".PowerOn_RetHome.Q) AND "QZ01RetEvt") AND NOT ("IZ02RetPos"),
                                         PT := T#5S);
   // 含义：条件 (((#MainStep.S2 AND NOT (#MainStep.S6)) AND "DB1042_Timer".DrillMemory) AND "DB1042_Timer".PowerOn_RetHome.Q) AND "DB1042_Timer".RetHome_Z02TimeOut.Q 成立时，将 TRUE 传送到 #MainStep.ErrEnd
   IF (((#MainStep.S2 AND NOT (#MainStep.S6)) AND "DB1042_Timer".DrillMemory) AND "DB1042_Timer".PowerOn_RetHome.Q) AND "DB1042_Timer".RetHome_Z02TimeOut.Q THEN
       #MainStep.ErrEnd := TRUE;
   END_IF;
   // 含义：条件 (((#MainStep.S2 AND NOT (#MainStep.S6)) AND "DB1042_Timer".DrillMemory) AND "DB1042_Timer".PowerOn_RetHome.Q) AND "DB1042_Timer".RetHome_Z02TimeOut.Q 成立时，将 TRUE 传送到 "DB1080_Component".Robot.Cmd.Auto.Stop
   IF (((#MainStep.S2 AND NOT (#MainStep.S6)) AND "DB1042_Timer".DrillMemory) AND "DB1042_Timer".PowerOn_RetHome.Q) AND "DB1042_Timer".RetHome_Z02TimeOut.Q THEN
       "DB1080_Component".Robot.Cmd.Auto.Stop := TRUE;
   END_IF;
   // 含义：条件 (((#MainStep.S2 AND NOT (#MainStep.S6)) AND "DB1042_Timer".DrillMemory) AND "DB1042_Timer".PowerOn_RetHome.Q) AND "DB1042_Timer".RetHome_Z02TimeOut.Q 成立时，将 TRUE 传送到 "DB1148_PromptBeeper".Public.RetHome_Z02RetTimeOut
   IF (((#MainStep.S2 AND NOT (#MainStep.S6)) AND "DB1042_Timer".DrillMemory) AND "DB1042_Timer".PowerOn_RetHome.Q) AND "DB1042_Timer".RetHome_Z02TimeOut.Q THEN
       "DB1148_PromptBeeper".Public.RetHome_Z02RetTimeOut := TRUE;
   END_IF;
   // 含义：条件 (((((#MainStep.S2 AND NOT (#MainStep.S6)) AND "DB1042_Timer".DrillMemory) AND "DB1042_Timer".PowerOn_RetHome.Q) AND "IZ02RetPos") AND "DB1081_ValveCall".ST01.Z02.RetPos) OR (((((#MainStep.S2 AND NOT (#MainStep.S6)) AND "DB1042_Timer".DrillMemory) AND "DB1042_Timer".PowerOn_RetHome.Q) AND "IZ02RetPos") AND "IZ02RetPos") 成立时，将 TRUE 传送到 #EdgeDetc.JUMP[0]
   IF (((((#MainStep.S2 AND NOT (#MainStep.S6)) AND "DB1042_Timer".DrillMemory) AND "DB1042_Timer".PowerOn_RetHome.Q) AND "IZ02RetPos") AND "DB1081_ValveCall".ST01.Z02.RetPos) OR (((((#MainStep.S2 AND NOT (#MainStep.S6)) AND "DB1042_Timer".DrillMemory) AND "DB1042_Timer".PowerOn_RetHome.Q) AND "IZ02RetPos") AND "IZ02RetPos") THEN
       #EdgeDetc.JUMP[0] := TRUE;
   END_IF;
   // 含义：条件 (((((#MainStep.S2 AND NOT (#MainStep.S6)) AND "DB1042_Timer".DrillMemory) AND "DB1042_Timer".PowerOn_RetHome.Q) AND "IZ02RetPos") AND "DB1081_ValveCall".ST01.Z02.RetPos) OR (((((#MainStep.S2 AND NOT (#MainStep.S6)) AND "DB1042_Timer".DrillMemory) AND "DB1042_Timer".PowerOn_RetHome.Q) AND "IZ02RetPos") AND "IZ02RetPos") 成立时，将 TRUE 传送到 "DB1080_Component".Robot.Cmd.Auto.ProgStart
   IF (((((#MainStep.S2 AND NOT (#MainStep.S6)) AND "DB1042_Timer".DrillMemory) AND "DB1042_Timer".PowerOn_RetHome.Q) AND "IZ02RetPos") AND "DB1081_ValveCall".ST01.Z02.RetPos) OR (((((#MainStep.S2 AND NOT (#MainStep.S6)) AND "DB1042_Timer".DrillMemory) AND "DB1042_Timer".PowerOn_RetHome.Q) AND "IZ02RetPos") AND "IZ02RetPos") THEN
       "DB1080_Component".Robot.Cmd.Auto.ProgStart := TRUE;
   END_IF;
   // 含义：条件 (((((#MainStep.S2 AND NOT (#MainStep.S6)) AND "DB1042_Timer".DrillMemory) AND "DB1042_Timer".PowerOn_RetHome.Q) AND "IZ02RetPos") AND "DB1081_ValveCall".ST01.Z02.RetPos) OR (((((#MainStep.S2 AND NOT (#MainStep.S6)) AND "DB1042_Timer".DrillMemory) AND "DB1042_Timer".PowerOn_RetHome.Q) AND "IZ02RetPos") AND "IZ02RetPos") 成立时，将 TRUE 传送到 "DB1080_Component".Robot.Cmd.Auto.GoHome
   IF (((((#MainStep.S2 AND NOT (#MainStep.S6)) AND "DB1042_Timer".DrillMemory) AND "DB1042_Timer".PowerOn_RetHome.Q) AND "IZ02RetPos") AND "DB1081_ValveCall".ST01.Z02.RetPos) OR (((((#MainStep.S2 AND NOT (#MainStep.S6)) AND "DB1042_Timer".DrillMemory) AND "DB1042_Timer".PowerOn_RetHome.Q) AND "IZ02RetPos") AND "IZ02RetPos") THEN
       "DB1080_Component".Robot.Cmd.Auto.GoHome := TRUE;
   END_IF;
   // 含义：条件 (((((#MainStep.S2 AND NOT (#MainStep.S6)) AND "DB1042_Timer".DrillMemory) AND "DB1042_Timer".PowerOn_RetHome.Q) AND "IZ02RetPos") AND "DB1081_ValveCall".ST01.Z02.RetPos) OR (((((#MainStep.S2 AND NOT (#MainStep.S6)) AND "DB1042_Timer".DrillMemory) AND "DB1042_Timer".PowerOn_RetHome.Q) AND "IZ02RetPos") AND "IZ02RetPos") 成立时，将 255 传送到 "DB1080_Component".Robot.CTRL_IN.ProgNo
   IF (((((#MainStep.S2 AND NOT (#MainStep.S6)) AND "DB1042_Timer".DrillMemory) AND "DB1042_Timer".PowerOn_RetHome.Q) AND "IZ02RetPos") AND "DB1081_ValveCall".ST01.Z02.RetPos) OR (((((#MainStep.S2 AND NOT (#MainStep.S6)) AND "DB1042_Timer".DrillMemory) AND "DB1042_Timer".PowerOn_RetHome.Q) AND "IZ02RetPos") AND "IZ02RetPos") THEN
       "DB1080_Component".Robot.CTRL_IN.ProgNo := 255;
   END_IF;
   // 含义：条件 #MainStep.S2 AND NOT (#MainStep.S6) 成立时，将 15 传送到 "DB1080_Component".Robot.CTRL_IN.RobotSpeed
   IF #MainStep.S2 AND NOT (#MainStep.S6) THEN
       "DB1080_Component".Robot.CTRL_IN.RobotSpeed := 15;
   END_IF;
   // 含义：条件 ((#MainStep.S2 AND #EdgeDetc.JUMP[0]) AND ("DB1900_Communication_PC".Recv.Current_2 < 0.5)) 成立时，将 TRUE 传送到 #MainStep.ErrEnd
   IF ((#MainStep.S2 AND #EdgeDetc.JUMP[0]) AND ("DB1900_Communication_PC".Recv.Current_2 < 0.5)) THEN
       #MainStep.ErrEnd := TRUE;
   END_IF;
   // 含义：条件 ((#MainStep.S2 AND #EdgeDetc.JUMP[0]) AND ("DB1900_Communication_PC".Recv.Current_2 < 0.5)) 成立时，将 TRUE 传送到 "DB1080_Component".Robot.Cmd.Auto.Stop
   IF ((#MainStep.S2 AND #EdgeDetc.JUMP[0]) AND ("DB1900_Communication_PC".Recv.Current_2 < 0.5)) THEN
       "DB1080_Component".Robot.Cmd.Auto.Stop := TRUE;
   END_IF;
   // 含义：条件 ((#MainStep.S2 AND #EdgeDetc.JUMP[0]) AND ("DB1900_Communication_PC".Recv.Current_2 < 0.5)) 成立时，将 TRUE 传送到 "DB1148_PromptBeeper".Public.RetHome_PowerOff
   IF ((#MainStep.S2 AND #EdgeDetc.JUMP[0]) AND ("DB1900_Communication_PC".Recv.Current_2 < 0.5)) THEN
       "DB1148_PromptBeeper".Public.RetHome_PowerOff := TRUE;
   END_IF;
   // 含义：条件 (#MainStep.S2 AND "DB1042_Timer".RetHomeHighCurrentOut.Q) OR (((#MainStep.S2 AND #EdgeDetc.JUMP[0]) AND ("DB1900_Communication_PC".Recv.Current_2 > "DB1900_Communication_PC".Para.CurrentMaxLimit))) 成立时，将 TRUE 传送到 #MainStep.ErrEnd
   IF (#MainStep.S2 AND "DB1042_Timer".RetHomeHighCurrentOut.Q) OR (((#MainStep.S2 AND #EdgeDetc.JUMP[0]) AND ("DB1900_Communication_PC".Recv.Current_2 > "DB1900_Communication_PC".Para.CurrentMaxLimit))) THEN
       #MainStep.ErrEnd := TRUE;
   END_IF;
   // 含义：条件 (#MainStep.S2 AND "DB1042_Timer".RetHomeHighCurrentOut.Q) OR (((#MainStep.S2 AND #EdgeDetc.JUMP[0]) AND ("DB1900_Communication_PC".Recv.Current_2 > "DB1900_Communication_PC".Para.CurrentMaxLimit))) 成立时，将 TRUE 传送到 "DB1080_Component".Robot.Cmd.Auto.Stop
   IF (#MainStep.S2 AND "DB1042_Timer".RetHomeHighCurrentOut.Q) OR (((#MainStep.S2 AND #EdgeDetc.JUMP[0]) AND ("DB1900_Communication_PC".Recv.Current_2 > "DB1900_Communication_PC".Para.CurrentMaxLimit))) THEN
       "DB1080_Component".Robot.Cmd.Auto.Stop := TRUE;
   END_IF;
   // 含义：条件 (#MainStep.S2 AND "DB1042_Timer".RetHomeHighCurrentOut.Q) OR (((#MainStep.S2 AND #EdgeDetc.JUMP[0]) AND ("DB1900_Communication_PC".Recv.Current_2 > "DB1900_Communication_PC".Para.CurrentMaxLimit))) 成立时，将 TRUE 传送到 "DB1148_PromptBeeper".Public.BitStuckErr_HighCurrent
   IF (#MainStep.S2 AND "DB1042_Timer".RetHomeHighCurrentOut.Q) OR (((#MainStep.S2 AND #EdgeDetc.JUMP[0]) AND ("DB1900_Communication_PC".Recv.Current_2 > "DB1900_Communication_PC".Para.CurrentMaxLimit))) THEN
       "DB1148_PromptBeeper".Public.BitStuckErr_HighCurrent := TRUE;
   END_IF;
   // 含义：将 (#MainStep.S2 AND "DB1080_Component".Robot.Status.HomePos) OR (#MainStep.S2 AND #MainStep.S6) 赋给 #MainStep.S6
   #MainStep.S6 := (#MainStep.S2 AND "DB1080_Component".Robot.Status.HomePos) OR (#MainStep.S2 AND #MainStep.S6);

   // ---------- 网络 8 ----------
   // 标题：枪电源
   // 含义：条件 #MainStep.S6 AND NOT (#MainStep.S8) 成立时，将 TRUE 传送到 "DB1081_ValveCall".ST01.Z05.RetAuto
   IF #MainStep.S6 AND NOT (#MainStep.S8) THEN
       "DB1081_ValveCall".ST01.Z05.RetAuto := TRUE;
   END_IF;
   // 含义：条件 #MainStep.S6 AND NOT (#MainStep.S8) 成立时，将 FALSE 传送到 #EdgeDetc.JUMP[0]
   IF #MainStep.S6 AND NOT (#MainStep.S8) THEN
       #EdgeDetc.JUMP[0] := FALSE;
   END_IF;
   // 含义：条件 #MainStep.S6 AND NOT (#MainStep.S8) 成立时，将 FALSE 传送到 "DB1042_Timer".DrillMemory
   IF #MainStep.S6 AND NOT (#MainStep.S8) THEN
       "DB1042_Timer".DrillMemory := FALSE;
   END_IF;
   // 含义：将 (#MainStep.S6 AND "DB1081_ValveCall".ST01.Z05.RetPos) OR (#MainStep.S6 AND #MainStep.S8) 赋给 #MainStep.S8
   #MainStep.S8 := (#MainStep.S6 AND "DB1081_ValveCall".ST01.Z05.RetPos) OR (#MainStep.S6 AND #MainStep.S8);

   // ---------- 网络 9 ----------
   // 标题：凿击三爪卡盘夹爪气缸
   // 含义：条件 (NOT (TRUE) AND NOT (#MainStep.S8)) AND NOT (#MainStep.S10) 成立时，将 TRUE 传送到 "DB1081_ValveCall".ST01.Z09.RetAuto
   IF (NOT (TRUE) AND NOT (#MainStep.S8)) AND NOT (#MainStep.S10) THEN
       "DB1081_ValveCall".ST01.Z09.RetAuto := TRUE;
   END_IF;
   // 含义：将 ((NOT (TRUE) AND NOT (#MainStep.S8)) AND "DB1081_ValveCall".ST01.Z09.RetPos) OR ((NOT (TRUE) AND NOT (#MainStep.S8)) AND TRUE) OR ((NOT (TRUE) AND NOT (#MainStep.S8)) AND NOT ("DB1900_Communication_PC".Para.ProduceMode3)) OR ((NOT (TRUE) AND NOT (#MainStep.S8)) AND #MainStep.S10) 赋给 #MainStep.S10
   #MainStep.S10 := ((NOT (TRUE) AND NOT (#MainStep.S8)) AND "DB1081_ValveCall".ST01.Z09.RetPos) OR ((NOT (TRUE) AND NOT (#MainStep.S8)) AND TRUE) OR ((NOT (TRUE) AND NOT (#MainStep.S8)) AND NOT ("DB1900_Communication_PC".Para.ProduceMode3)) OR ((NOT (TRUE) AND NOT (#MainStep.S8)) AND #MainStep.S10);

   // ---------- 网络 10 ----------
   // 标题：推力气缸
   // 含义：条件 (#MainStep.S8 OR #MainStep.S10) AND NOT (#MainStep.S13) 成立时，将 TRUE 传送到 "DB1081_ValveCall".ST01.Z01.ExtAuto
   IF (#MainStep.S8 OR #MainStep.S10) AND NOT (#MainStep.S13) THEN
       "DB1081_ValveCall".ST01.Z01.ExtAuto := TRUE;
   END_IF;
   // 含义：条件 (#MainStep.S8 OR #MainStep.S10) AND NOT (#MainStep.S13) 成立时，将 TRUE 传送到 "DB1081_ValveCall".ST01.Z02.VentValveAuto
   IF (#MainStep.S8 OR #MainStep.S10) AND NOT (#MainStep.S13) THEN
       "DB1081_ValveCall".ST01.Z02.VentValveAuto := TRUE;
   END_IF;
   // 含义：条件 (#MainStep.S8 OR #MainStep.S10) AND NOT (#MainStep.S13) 成立时，将 TRUE 传送到 "DB1081_ValveCall".ST01.Z05.RetAuto
   IF (#MainStep.S8 OR #MainStep.S10) AND NOT (#MainStep.S13) THEN
       "DB1081_ValveCall".ST01.Z05.RetAuto := TRUE;
   END_IF;
   // 含义：条件 (#MainStep.S8 OR #MainStep.S10) AND NOT (#MainStep.S13) 成立时，将 TRUE 传送到 "DB1081_ValveCall".ST01.Z08.RetAuto
   IF (#MainStep.S8 OR #MainStep.S10) AND NOT (#MainStep.S13) THEN
       "DB1081_ValveCall".ST01.Z08.RetAuto := TRUE;
   END_IF;
   // 含义：条件 (#MainStep.S8 OR #MainStep.S10) AND NOT (#MainStep.S13) 成立时，将 FALSE 传送到 "DB1080_Component".Robot.Cmd.Auto.GoHome
   IF (#MainStep.S8 OR #MainStep.S10) AND NOT (#MainStep.S13) THEN
       "DB1080_Component".Robot.Cmd.Auto.GoHome := FALSE;
   END_IF;
   // 含义：条件 ((((#MainStep.S8 OR #MainStep.S10) AND NOT (#MainStep.S13)) AND ("DB720_KuKa_MainCtrl".CmdOut.gi_ToolTypeNo = 13))) AND TRUE 成立时，将 FALSE 传送到 "QCamCoverExt"
   IF ((((#MainStep.S8 OR #MainStep.S10) AND NOT (#MainStep.S13)) AND ("DB720_KuKa_MainCtrl".CmdOut.gi_ToolTypeNo = 13))) AND TRUE THEN
       "QCamCoverExt" := FALSE;
   END_IF;
   // 含义：条件 ((((#MainStep.S8 OR #MainStep.S10) AND NOT (#MainStep.S13)) AND ("DB720_KuKa_MainCtrl".CmdOut.gi_ToolTypeNo = 13))) AND TRUE 成立时，将 TRUE 传送到 "QCamCoverRet"
   IF ((((#MainStep.S8 OR #MainStep.S10) AND NOT (#MainStep.S13)) AND ("DB720_KuKa_MainCtrl".CmdOut.gi_ToolTypeNo = 13))) AND TRUE THEN
       "QCamCoverRet" := TRUE;
   END_IF;
   // 含义：条件 (#MainStep.S8 OR #MainStep.S10) AND NOT (#MainStep.S13) 成立时，将 0.3 传送到 "DB1080_Component".Aux.Pressure
   IF (#MainStep.S8 OR #MainStep.S10) AND NOT (#MainStep.S13) THEN
       "DB1080_Component".Aux.Pressure := 0.3;
   END_IF;
   // 含义：将 ((((#MainStep.S8 OR #MainStep.S10) AND "DB1081_ValveCall".ST01.Z01.ExtPos) AND "IZ02ExtPos") AND "DB1081_ValveCall".ST01.Z05.RetPos) OR ((#MainStep.S8 OR #MainStep.S10) AND #MainStep.S13) 赋给 #MainStep.S13
   #MainStep.S13 := ((((#MainStep.S8 OR #MainStep.S10) AND "DB1081_ValveCall".ST01.Z01.ExtPos) AND "IZ02ExtPos") AND "DB1081_ValveCall".ST01.Z05.RetPos) OR ((#MainStep.S8 OR #MainStep.S10) AND #MainStep.S13);

   // ---------- 网络 11 ----------
   // 标题：右防尘盖夹紧缸
   // 含义：条件 (#MainStep.S13 AND NOT (#MainStep.S17)) AND "DB720_KuKa_MainCtrl".Aux.AStation_ToolAtPosT.Q 成立时，将 TRUE 传送到 "DB1081_ValveCall".ST01.Z03.RetAuto
   IF (#MainStep.S13 AND NOT (#MainStep.S17)) AND "DB720_KuKa_MainCtrl".Aux.AStation_ToolAtPosT.Q THEN
       "DB1081_ValveCall".ST01.Z03.RetAuto := TRUE;
   END_IF;
   // 含义：条件 (#MainStep.S13 AND NOT (#MainStep.S17)) AND "DB720_KuKa_MainCtrl".Aux.BStation_ToolAtPosT.Q 成立时，将 TRUE 传送到 "DB1081_ValveCall".ST01.Z04.RetAuto
   IF (#MainStep.S13 AND NOT (#MainStep.S17)) AND "DB720_KuKa_MainCtrl".Aux.BStation_ToolAtPosT.Q THEN
       "DB1081_ValveCall".ST01.Z04.RetAuto := TRUE;
   END_IF;
   // 含义：将 (((#MainStep.S13 AND "DB1081_ValveCall".ST01.Z03.RetPos) OR (#MainStep.S13 AND NOT ("DB720_KuKa_MainCtrl".Aux.AStation_ToolAtPosT.Q))) AND "DB1081_ValveCall".ST01.Z04.RetPos) OR (((#MainStep.S13 AND "DB1081_ValveCall".ST01.Z03.RetPos) OR (#MainStep.S13 AND NOT ("DB720_KuKa_MainCtrl".Aux.AStation_ToolAtPosT.Q))) AND NOT ("DB720_KuKa_MainCtrl".Aux.BStation_ToolAtPosT.Q)) OR (#MainStep.S13 AND #MainStep.S17) 赋给 #MainStep.S17
   #MainStep.S17 := (((#MainStep.S13 AND "DB1081_ValveCall".ST01.Z03.RetPos) OR (#MainStep.S13 AND NOT ("DB720_KuKa_MainCtrl".Aux.AStation_ToolAtPosT.Q))) AND "DB1081_ValveCall".ST01.Z04.RetPos) OR (((#MainStep.S13 AND "DB1081_ValveCall".ST01.Z03.RetPos) OR (#MainStep.S13 AND NOT ("DB720_KuKa_MainCtrl".Aux.AStation_ToolAtPosT.Q))) AND NOT ("DB720_KuKa_MainCtrl".Aux.BStation_ToolAtPosT.Q)) OR (#MainStep.S13 AND #MainStep.S17);

   // ---------- 网络 12 ----------
   // 含义：将 #MainStep.S17 OR #MainStep.ErrEnd 赋给 #MainStep.End
   #MainStep.End := #MainStep.S17 OR #MainStep.ErrEnd;

   // ---------- 网络 13 ----------
   // （空白网络）
END_FUNCTION_BLOCK

// folder: 004_AutoStep

FUNCTION_BLOCK "FB720_KuKa_MainCtrl"   // FB720, SCL
{ S7_Optimized_Access := 'TRUE' }
// ============================================================
//  Block: FB720_KuKa_MainCtrl
//  ============================================================
//  编号：FB720
//  原始语言：LAD（规则翻译为 SCL）
//  含义：Thrust Cylinder in Extend Position When Changing Tools, Programmed  By WXY 20230307,
   VAR
      CmdOut : Struct   // 总共56个Byte,自定义输入状态
         di_ChgGrp_Ack : Bool;   // 换爪完成确认
         di_HorDril_Ack : Bool;   // 水平钻入开始确认
         di_DiamondVib_Ack : Bool;   // 水钻岩芯敲击完成确认
         di_DownDril_Ack : Bool;   // 向下钻入开始确认
         di_ChkScrew_Ack : Bool;   // 检查钻头完成确认
         di_Drilling_Ack : Bool;   // 开始钻孔确认
         di_StopDril_Ack : Bool;   // 停止钻孔确认
         di_Front_Sig : Bool;   // 推力气缸前端
         di_StopDrill_End : Bool;   // 请求打孔结束
         di_Middle_Sig : Bool;   // 推力气缸中间
         di_Stop_Sig : Bool;   // 推力气缸停止
         di_DiamondDetc_Ack : Bool;   // 水钻岩芯检测完成确认
         di_Gouge_Ack : Bool;   // 凿击完成确认
         di_ToolPos : Bool;   // 工装有无
         di_TouchPos : Bool;   // 接触到水泥确认，用于机器人计算进给
         di_VchiselTime_End : Bool;   // 凿击时间结束
         di_VchiselCamera_End : Bool;   // 视觉凿击相机拍照流程结束
         di_ChiselCylinderRet : Bool;   // 凿击退出辅助气缸缩回
         di_ChiselRobotRet : Bool;   // 凿击机器人退出
         di_DownChiselMode : Bool;   // 向下凿击模式
         di_PushCylOK_Sig : Bool;   // 凿击推力气缸推出到位
         di_FTCalib_End : Bool;   // 力控校准完毕
         di_FTAction_Cmd : Bool;   // 力控调整指令
         di_NotDectceDiamond : Bool;   // 不检测水钻岩芯
         gi_ToolPosNo : Byte;   // 夹具位置号
         gi_LayerNum : Byte;   // 凿击层数
         gi_VChiselCamShotArea : Byte;   // 水平视觉凿击拍照位置
         gi_OffSetX : DWord;   // X方向偏移值
         gi_OffSetY : DWord;   // Y方向偏移值
         gi_OffSetZ : DWord;   // Z方向偏移值
         gi_Depth : DWord;   // 钻入深度
         gi_ScrewLength : DWord;   // 批头长度
         gi_Angle : DWord;   // 角度
         gi_Width : DWord;   // 凿钻间距
         gi_OffSetA : DWord;   // 静态变量
         gi_OffSetB : DWord;   // 静态变量
         gi_OffSetC : DWord;   // 静态变量
         gi_DownSlabHeight : DWord;   // 向下水泥块厚度
         gi_ToolTypeNo : Byte;   // 静态变量
         gi_Spare : Byte;   // 静态变量
         SP : Array[1..4] of Byte;   // 静态变量
      END_STRUCT;
      ATCmdOut : Array[8..63] of Byte;   // To Robot
      StatusIn : Struct   // 总共56个Byte,自定义输出命令
         do_ChgGrp_Act : Bool;   // 换爪运行中
         do_HorDril_Act : Bool;   // 水平方向钻入运行中
         do_UpDril_Act : Bool;   // 向上方向钻入运行中
         do_DownDril_Act : Bool;   // 向下方向钻入运行中
         do_ChkScrew_Act : Bool;   // 检查钻头运行中
         do_Diamond_Act : Bool;   // 水钻岩芯敲击运行中
         do_DrillReady_Act : Bool;   // 转孔就位
         do_Gouge_Act : Bool;   // 凿击运行中
         do_DiamondDetc_Pos : Bool;   // 水钻岩芯检测位置
         do_CameraPos_Ready : Bool;   // 视觉相机在拍照位
         do_RobotPry_End : Bool;   // 机器人摆动结束(视觉凿击)
         do_ChiselCylinderExt : Bool;   // 凿击模式下IN点气缸推出
         do_FixStationToHome : Bool;   // 机器人在夹具位置回原点
         do_FTCalibPos : Bool;   // 机器人到达力控校准点
         do_FTAction_Rcv : Bool;   // 机器人接收到力控调整指令
         do_DownDrilApp_Pos : Bool;   // 向下钻孔接近位置
         do_ChgGrp_Pos : Bool;   // 换爪位置
         do_HorDril_Pos : Bool;   // 水平方向钻入位置
         do_JDiamond_MidPos : Bool;   // 水钻岩芯过渡位置
         do_DownDril_Pos : Bool;   // 向下方向钻入位置
         do_ChkScrew_Pos : Bool;   // 检查钻头位置
         do_ReqDrilling : Bool;   // 请求钻孔
         do_ReqStopDril : Bool;   // 请求停止钻孔
         do_DiamondVib_Pos : Bool;   // 水钻岩芯敲击位置
         do_Gouge_Pos : Bool;   // 凿击位置
         do_DrilEnd_Pos : Bool;   // End点位置
         do_ChiselPry : Bool;   // 凿击摆动
         SPARE3 : Bool;   // 静态变量
         SPARE4 : Bool;   // 静态变量
         SPARE5 : Bool;   // 静态变量
         SPARE6 : Bool;   // 静态变量
         SPARE7 : Bool;   // 静态变量
         do_ChgGrp_Don : Bool;   // 换爪完成
         do_HorDril_Don : Bool;   // 水平方向钻入完成
         do_UpDril_Don : Bool;   // 向上方向钻入完成
         do_DownDril_Don : Bool;   // 向下方向钻入完成
         do_ChkScrew_Don : Bool;   // 检查钻头完成
         do_Diamond_Don : Bool;   // 水钻岩芯去除完成
         do_Gouge_Don : Bool;   // 凿击完成
         do_Gouge_Don1 : Bool;   // 静态变量
         Static_8 : Byte;   // 静态变量
         do_NotInGripLib_Area : Bool;   // 不在夹具库范围
         do_NotInHor_Area : Bool;   // 不在水平钻孔范围
         do_NotInGripLib_Area_1 : Bool;   // 不在向上钻孔范围
         do_NotInGripLib_Area_2 : Bool;   // 不在向下钻孔范围
         Static_1 : Byte;   // 静态变量
         Static_2 : Byte;   // 静态变量
         Static_3 : Byte;   // 静态变量
         go_X : Real;   // 静态变量
         go_Y : Real;   // 静态变量
         go_Z : Real;   // 静态变量
         SP : Array[1..33] of Byte;   // 静态变量
      END_STRUCT;
      AtStatusIn : Array[8..63] of Byte;   // To Plc
      Ctrl_Out : Struct   // 静态变量
         RobotAction : DInt;   // 机器人调用流程已启用
      END_STRUCT;
      AtCtrl_Out : Struct   // 静态变量
         RobotAction : Struct   // 静态变量
            SP : Int;   // 静态变量
            GetTray : Bool;   // 静态变量
            PutTray : Bool;   // 静态变量
            GetPed : Bool;   // 静态变量
            PutPed : Bool;   // 静态变量
            PutAssembly : Bool;   // 静态变量
            GetAssembly : Bool;   // 静态变量
            PutTest : Bool;   // 静态变量
            GetTest : Bool;   // 静态变量
            PutCirclip : Bool;   // 静态变量
            GetGearBox : Bool;   // 静态变量
            PutProduct : Bool;   // 静态变量
            GetTool : Bool;   // 静态变量
            PutTool : Bool;   // 静态变量
         END_STRUCT;
      END_STRUCT;
      CheckBit : Struct   // 检查批头
         Busy : Bool;   // 静态变量
         StartCmd : Bool;   // 静态变量
         OKToStart : Bool;   // 静态变量
         TaskDone : Bool;   // 静态变量
         StepStart : Bool;   // 静态变量
         StepEnd : Bool;   // 静态变量
         ErrEnd : Bool;   // 静态变量
         ByPass : Bool;   // 静态变量
         TaskIO : Bool;   // 静态变量
         TaskNIO : Bool;   // 静态变量
         S1 : Bool;   // 静态变量
         S2 : Bool;   // 静态变量
         S3 : Bool;   // 静态变量
         S4 : Bool;   // 静态变量
         S5 : Bool;   // 静态变量
         S6 : Bool;   // 静态变量
         S7 : Bool;   // 静态变量
         S8 : Bool;   // 静态变量
         S9 : Bool;   // 静态变量
         S10 : Bool;   // 静态变量
         S11 : Bool;   // 静态变量
         S12 : Bool;   // 静态变量
         S13 : Bool;   // 静态变量
         S14 : Bool;   // 静态变量
         S15 : Bool;   // 静态变量
         S16 : Bool;   // 静态变量
         S17 : Bool;   // 静态变量
         S18 : Bool;   // 静态变量
         S19 : Bool;   // 静态变量
         S20 : Bool;   // 静态变量
         S21 : Bool;   // 静态变量
         S22 : Bool;   // 静态变量
         S23 : Bool;   // 静态变量
         S24 : Bool;   // 静态变量
         S25 : Bool;   // 静态变量
         S26 : Bool;   // 静态变量
         S27 : Bool;   // 静态变量
         S28 : Bool;   // 静态变量
         S29 : Bool;   // 静态变量
         S30 : Bool;   // 静态变量
         S31 : Bool;   // 静态变量
         S32 : Bool;   // 静态变量
         S33 : Bool;   // 静态变量
         S34 : Bool;   // 静态变量
         S35 : Bool;   // 静态变量
         S36 : Bool;   // 静态变量
         S37 : Bool;   // 静态变量
         S38 : Bool;   // 静态变量
         S39 : Bool;   // 静态变量
         S40 : Bool;   // 静态变量
         S41 : Bool;   // 静态变量
         S42 : Bool;   // 静态变量
         S43 : Bool;   // 静态变量
         S44 : Bool;   // 静态变量
         S45 : Bool;   // 静态变量
         S46 : Bool;   // 静态变量
         S47 : Bool;   // 静态变量
         S48 : Bool;   // 静态变量
         S49 : Bool;   // 静态变量
         S50 : Bool;   // 静态变量
         S51 : Bool;   // 静态变量
         S52 : Bool;   // 静态变量
         S53 : Bool;   // 静态变量
         S54 : Bool;   // 静态变量
         S55 : Bool;   // 静态变量
         S56 : Bool;   // 静态变量
         S57 : Bool;   // 静态变量
         S58 : Bool;   // 静态变量
         S59 : Bool;   // 静态变量
         S60 : Bool;   // 静态变量
         S61 : Bool;   // 静态变量
         S62 : Bool;   // 静态变量
         S63 : Bool;   // 静态变量
         S64 : Bool;   // 静态变量
         S65 : Bool;   // 静态变量
         S66 : Bool;   // 静态变量
         S67 : Bool;   // 静态变量
      END_STRUCT;
      ChangeTool : Struct   // 换爪
         Busy : Bool;   // 静态变量
         StartCmd : Bool;   // 静态变量
         OKToStart : Bool;   // 静态变量
         TaskDone : Bool;   // 静态变量
         StepStart : Bool;   // 静态变量
         StepEnd : Bool;   // 静态变量
         ErrEnd : Bool;   // 静态变量
         ByPass : Bool;   // 静态变量
         TaskIO : Bool;   // 静态变量
         TaskNIO : Bool;   // 静态变量
         S1 : Bool;   // 静态变量
         S2 : Bool;   // 静态变量
         S3 : Bool;   // 静态变量
         S4 : Bool;   // 静态变量
         S5 : Bool;   // 静态变量
         S6 : Bool;   // 静态变量
         S7 : Bool;   // 静态变量
         S8 : Bool;   // 静态变量
         S9 : Bool;   // 静态变量
         S10 : Bool;   // 静态变量
         S11 : Bool;   // 静态变量
         S12 : Bool;   // 静态变量
         S13 : Bool;   // 静态变量
         S14 : Bool;   // 静态变量
         S15 : Bool;   // 静态变量
         S16 : Bool;   // 静态变量
         S17 : Bool;   // 静态变量
         S18 : Bool;   // 静态变量
         S19 : Bool;   // 静态变量
         S20 : Bool;   // 静态变量
         S21 : Bool;   // 静态变量
         S22 : Bool;   // 静态变量
         S23 : Bool;   // 静态变量
         S24 : Bool;   // 静态变量
         S25 : Bool;   // 静态变量
         S26 : Bool;   // 静态变量
         S27 : Bool;   // 静态变量
         S28 : Bool;   // 静态变量
         S29 : Bool;   // 静态变量
         S30 : Bool;   // 静态变量
         S31 : Bool;   // 静态变量
         S32 : Bool;   // 静态变量
         S33 : Bool;   // 静态变量
         S34 : Bool;   // 静态变量
         S35 : Bool;   // 静态变量
         S36 : Bool;   // 静态变量
         S37 : Bool;   // 静态变量
         S38 : Bool;   // 静态变量
         S39 : Bool;   // 静态变量
         S40 : Bool;   // 静态变量
         S41 : Bool;   // 静态变量
         S42 : Bool;   // 静态变量
         S43 : Bool;   // 静态变量
         S44 : Bool;   // 静态变量
         S45 : Bool;   // 静态变量
         S46 : Bool;   // 静态变量
         S47 : Bool;   // 静态变量
         S48 : Bool;   // 静态变量
         S49 : Bool;   // 静态变量
         S50 : Bool;   // 静态变量
         S51 : Bool;   // 静态变量
         S52 : Bool;   // 静态变量
         S53 : Bool;   // 静态变量
         S54 : Bool;   // 静态变量
         S55 : Bool;   // 静态变量
         S56 : Bool;   // 静态变量
         S57 : Bool;   // 静态变量
         S58 : Bool;   // 静态变量
         S59 : Bool;   // 静态变量
         S60 : Bool;   // 静态变量
         S61 : Bool;   // 静态变量
         S62 : Bool;   // 静态变量
         S63 : Bool;   // 静态变量
         S64 : Bool;   // 静态变量
         S65 : Bool;   // 静态变量
         S66 : Bool;   // 静态变量
         S67 : Bool;   // 静态变量
      END_STRUCT;
      Aux : Struct   // 静态变量
         ToolAtPos : Bool;   // 机器人夹具在位置
         ToolRight : Bool;   // 静态变量
         BStation_oolAtPos : Bool;   // 右侧夹具在位置
         AStation_ToolAtPos : Bool;   // 左侧夹具在位置
         ToolAtPosTimer : IEC_TIMER;   // 夹具在位检测延时
         ToolNotAtPosTimer : IEC_TIMER;   // 夹具不在位检测延时
         AStation_ToolAtPosT : IEC_TIMER;   // 静态变量
         BStation_ToolAtPosT : IEC_TIMER;   // 静态变量
         ZeroPos : Real;   // 零点推力压缩长度
         OffSetY : Int;   // 静态变量
         OffSetYMid : DInt;   // 静态变量
         OffSetZ : Int;   // 静态变量
         OffSetZMid : DInt;   // 静态变量
         DrillDepth : Int;   // 静态变量
         DrillDepthMid : DInt;   // 静态变量
         ScrLen : Real;   // 静态变量
         ScrLen_Mid0 : DInt;   // 静态变量
         ScrLen_Mid1 : Real;   // 静态变量
         XZeroPos : Real;   // 水平钻孔开始X坐标
         ZZeroPos : Real;   // 水平钻孔开始Z坐标
         CurrentRobPos : Real;   // 当前机器人X坐标
         go_X : Real;   // 静态变量
         go_Z : Real;   // 静态变量
         MidPos_X : DInt;   // 静态变量
         MidPos_Z : DInt;   // 静态变量
         RobotSpeed : DInt;   // 静态变量
         LastToolPosNo : Int;   // 静态变量
         CheckNo : Int;   // 1水平2.向上3.向下
         PressureMid : Real;   // 静态变量
         Pressure : Real;   // 静态变量
         ForceNum : Int;   // 力数据编号
         DownSlabHeight : Int;   // 静态变量
      END_STRUCT;
      EdgeDetc : Struct   // 静态变量
         Pulse : Array[0..15] of Bool;   // 静态变量
      END_STRUCT;
      PT : Time;   // 静态变量
      ET : Time;   // 静态变量
      IN : Bool;   // 静态变量
      Q : Bool;   // 静态变量
   END_VAR
   VAR_TEMP
      T_Ret : Int;   // 临时变量
   END_VAR
   VAR CONSTANT
      Calculate_RobotProg_K : Int := 20;
   END_VAR
BEGIN

   // ---------- 网络 1 ----------
   // 标题：将用于自定义命令传入机器人
   // 含义：将 #ATCmdOut 赋给 "DB1080_Component".Robot.Bus_Out_Data.UserDefineRobIn
   "DB1080_Component".Robot.Bus_Out_Data.UserDefineRobIn := #ATCmdOut;
   // 含义：条件 NOT ("AllMode_M") 成立时，将 FALSE 传送到 "DB1148_PromptBeeper".Public.DrillDepthErr
   IF NOT ("AllMode_M") THEN
       "DB1148_PromptBeeper".Public.DrillDepthErr := FALSE;
   END_IF;
   // 含义：条件 NOT ("AllMode_M") 成立时，将 FALSE 传送到 "DB1148_PromptBeeper".Public.DrillTimeOut
   IF NOT ("AllMode_M") THEN
       "DB1148_PromptBeeper".Public.DrillTimeOut := FALSE;
   END_IF;
   // 含义：条件 NOT ("AllMode_M") 成立时，将 FALSE 传送到 "DB1148_PromptBeeper".Public.CurrentLowTimeOut
   IF NOT ("AllMode_M") THEN
       "DB1148_PromptBeeper".Public.CurrentLowTimeOut := FALSE;
   END_IF;
   // 含义：条件 NOT ("AllMode_M") 成立时，将 FALSE 传送到 "DB1148_PromptBeeper".Public.CurrentHighTimeOut
   IF NOT ("AllMode_M") THEN
       "DB1148_PromptBeeper".Public.CurrentHighTimeOut := FALSE;
   END_IF;
   // 含义：将 "DB1060_AutoStep".HorDrillAutoStep.HorDrillStep.StopDrill_Ack OR "DB1060_AutoStep".HorDrillAutoStep.HorDrillStep.GougeStopDrill_Ack OR "DB1060_AutoStep".DownDrillAutoStep.DownDrillStep.StopDrill_Ack 赋给 #CmdOut.di_StopDril_Ack
   #CmdOut.di_StopDril_Ack := "DB1060_AutoStep".HorDrillAutoStep.HorDrillStep.StopDrill_Ack OR "DB1060_AutoStep".HorDrillAutoStep.HorDrillStep.GougeStopDrill_Ack OR "DB1060_AutoStep".DownDrillAutoStep.DownDrillStep.StopDrill_Ack;
   // 含义：将 "DB1060_AutoStep".HorDrillAutoStep.HorDrillStep.StopDrill_End OR "DB1060_AutoStep".HorDrillAutoStep.HorDrillStep.GougeStopDrill_End OR "DB1060_AutoStep".DownDrillAutoStep.DownDrillStep.StopDrill_End OR "IZ02RetPos" OR ("DB1080_Component".ClinyderPos.Ctrl_Out.Cur_Val_Out > 82.0) 赋给 #CmdOut.di_StopDrill_End
   #CmdOut.di_StopDrill_End := "DB1060_AutoStep".HorDrillAutoStep.HorDrillStep.StopDrill_End OR "DB1060_AutoStep".HorDrillAutoStep.HorDrillStep.GougeStopDrill_End OR "DB1060_AutoStep".DownDrillAutoStep.DownDrillStep.StopDrill_End OR "IZ02RetPos" OR ("DB1080_Component".ClinyderPos.Ctrl_Out.Cur_Val_Out > 82.0);

   // ---------- 网络 2 ----------
   // 标题：向下水泥块厚度不在限制范围内(370-430)
   // 含义：条件 "ManMode_M" 成立时，将 ("DB1900_Communication_PC".Recv.DownSlabHeight - 0) 传送到 #Aux.DownSlabHeight
   IF "ManMode_M" THEN
       #Aux.DownSlabHeight := ("DB1900_Communication_PC".Recv.DownSlabHeight - 0);
   END_IF;
   // InRange uid=42 resolved
   // 含义：将 SWAP(#Aux.DownSlabHeight) 赋给 #CmdOut.gi_DownSlabHeight
   #CmdOut.gi_DownSlabHeight := SWAP(#Aux.DownSlabHeight);
   // OutRange uid=44 resolved
   // 含义：将 TRUE 赋给 "DB1060_AutoStep".DownDrillAutoStep.DownDrillStep.ErrEnd
   "DB1060_AutoStep".DownDrillAutoStep.DownDrillStep.ErrEnd := TRUE;
   // 含义：将 TRUE 赋给 "DB1148_PromptBeeper".Public.DownHeightErr
   "DB1148_PromptBeeper".Public.DownHeightErr := TRUE;
   // 含义：条件 "ManMode_M" AND "ErrRst_M" 成立时，将 FALSE 传送到 "DB1148_PromptBeeper".Public.DownHeightErr
   IF "ManMode_M" AND "ErrRst_M" THEN
       "DB1148_PromptBeeper".Public.DownHeightErr := FALSE;
   END_IF;

   // ---------- 网络 3 ----------
   // 标题：信号夹具ID号错误，请检查夹具！
   // 含义：调用定时器实例 #Aux.ToolAtPosTimer.TON
   #Aux.ToolAtPosTimer.TON(IN := "IToolAtPos",
                           PT := T#100ms);
   // 含义：调用定时器实例 #Aux.ToolNotAtPosTimer.TON
   #Aux.ToolNotAtPosTimer.TON(IN := NOT ("IToolAtPos"),
                              PT := T#100ms);
   // 含义：当 "IToolAtPos" 为 TRUE 时置位 #Aux.ToolAtPos，否则复位（触点→线圈）
   IF "IToolAtPos" THEN
       #Aux.ToolAtPos := TRUE;
   ELSE
       #Aux.ToolAtPos := FALSE;
   END_IF;
   // 含义：当 "IToolAtPos" 为 TRUE 时置位 #CmdOut.di_ToolPos，否则复位（触点→线圈）
   IF "IToolAtPos" THEN
       #CmdOut.di_ToolPos := TRUE;
   ELSE
       #CmdOut.di_ToolPos := FALSE;
   END_IF;
   // 含义：将 (("DB1900_Communication_PC".Para.IOFixtureNo = "DB1080_Component".IOFixtureIID.TP_CurFixtureID) AND ("DB1900_Communication_PC".Para.PowerFixtureNo = "DB1080_Component".PowerFixtureID.TP_CurFixtureID)) 赋给 #Aux.ToolRight
   #Aux.ToolRight := (("DB1900_Communication_PC".Para.IOFixtureNo = "DB1080_Component".IOFixtureIID.TP_CurFixtureID) AND ("DB1900_Communication_PC".Para.PowerFixtureNo = "DB1080_Component".PowerFixtureID.TP_CurFixtureID));
   // 含义：调用定时器实例 #Aux.AStation_ToolAtPosT.TON
   #Aux.AStation_ToolAtPosT.TON(IN := "AStation_ToolOn1" AND "AStation_ToolOn2",
                                PT := T#100ms);
   // 含义：调用定时器实例 #Aux.BStation_ToolAtPosT.TON
   #Aux.BStation_ToolAtPosT.TON(IN := "BStation_ToolOn1" AND "BStation_ToolOn2",
                                PT := T#100ms);
   // 含义：将 ((((("DB1080_Component".ClinyderPos.Ctrl_Out.Cur_Val_Out > 5.0) AND ("DB1080_Component".ClinyderPos.Ctrl_Out.Cur_Val_Out < 15.0))) AND ("DB1900_Communication_PC".Recv.ChooseProgNo = 4))) OR (((("DB1080_Component".ClinyderPos.Ctrl_Out.Cur_Val_Out > 5.0) AND ("DB1080_Component".ClinyderPos.Ctrl_Out.Cur_Val_Out < 15.0))) AND "ASMMode_M") OR (((((("DB1080_Component".ClinyderPos.Ctrl_Out.Cur_Val_Out > 60.0) AND ("DB1080_Component".ClinyderPos.Ctrl_Out.Cur_Val_Out < 80.0))) AND NOT ("ASMMode_M")) AND ("DB1900_Communication_PC".Recv.ChooseProgNo = 5))) 赋给 #CmdOut.di_Front_Sig
   #CmdOut.di_Front_Sig := ((((("DB1080_Component".ClinyderPos.Ctrl_Out.Cur_Val_Out > 5.0) AND ("DB1080_Component".ClinyderPos.Ctrl_Out.Cur_Val_Out < 15.0))) AND ("DB1900_Communication_PC".Recv.ChooseProgNo = 4))) OR (((("DB1080_Component".ClinyderPos.Ctrl_Out.Cur_Val_Out > 5.0) AND ("DB1080_Component".ClinyderPos.Ctrl_Out.Cur_Val_Out < 15.0))) AND "ASMMode_M") OR (((((("DB1080_Component".ClinyderPos.Ctrl_Out.Cur_Val_Out > 60.0) AND ("DB1080_Component".ClinyderPos.Ctrl_Out.Cur_Val_Out < 80.0))) AND NOT ("ASMMode_M")) AND ("DB1900_Communication_PC".Recv.ChooseProgNo = 5)));
   // 含义：将 ((("DB1080_Component".ClinyderPos.Ctrl_Out.Cur_Val_Out > 40.0) AND ("DB1080_Component".ClinyderPos.Ctrl_Out.Cur_Val_Out < 50.0))) AND NOT (TRUE) 赋给 #CmdOut.di_Middle_Sig
   #CmdOut.di_Middle_Sig := ((("DB1080_Component".ClinyderPos.Ctrl_Out.Cur_Val_Out > 40.0) AND ("DB1080_Component".ClinyderPos.Ctrl_Out.Cur_Val_Out < 50.0))) AND NOT (TRUE);
   // 含义：将 "DB1060_AutoStep".DownDrillAutoStep.DownDrillStep.StepStart OR "DB1060_AutoStep".HorDrillAutoStep.HorDrillStep.StepStart 赋给 "DB1900_Communication_PC".Send.RobotDrill
   "DB1900_Communication_PC".Send.RobotDrill := "DB1060_AutoStep".DownDrillAutoStep.DownDrillStep.StepStart OR "DB1060_AutoStep".HorDrillAutoStep.HorDrillStep.StepStart;

   // ---------- 网络 4 ----------
   // 标题：推力缸初始位置不正确！
   // 含义：将 (((("DB1060_AutoStep".HorDrillAutoStep.HorDrillStep.S10 AND NOT ("DB1060_AutoStep".HorDrillAutoStep.HorDrillStep.S12)) AND NOT ("DB1900_Communication_PC".Para.ProduceMode3)) OR (("DB1060_AutoStep".DownDrillAutoStep.DownDrillStep.S10 AND NOT ("DB1060_AutoStep".DownDrillAutoStep.DownDrillStep.S12)) AND NOT ("DB1900_Communication_PC".Para.ProduceMode3))) AND ("DB1080_Component".ClinyderPos.Ctrl_Out.Cur_Val_Out > 3.0)) 赋给 "DB1148_PromptBeeper".Public.Z01StartPosErr
   "DB1148_PromptBeeper".Public.Z01StartPosErr := (((("DB1060_AutoStep".HorDrillAutoStep.HorDrillStep.S10 AND NOT ("DB1060_AutoStep".HorDrillAutoStep.HorDrillStep.S12)) AND NOT ("DB1900_Communication_PC".Para.ProduceMode3)) OR (("DB1060_AutoStep".DownDrillAutoStep.DownDrillStep.S10 AND NOT ("DB1060_AutoStep".DownDrillAutoStep.DownDrillStep.S12)) AND NOT ("DB1900_Communication_PC".Para.ProduceMode3))) AND ("DB1080_Component".ClinyderPos.Ctrl_Out.Cur_Val_Out > 3.0));

   // ---------- 网络 5 ----------
   // 标题：*************************机器人坐标数据传递 深度计算*********************************
   // 含义：将 SWAP(#StatusIn.go_X) 赋给 #Aux.MidPos_X
   #Aux.MidPos_X := SWAP(#StatusIn.go_X);
   // 含义：将 #Aux.MidPos_X; (* Convert → Real *) 赋给 #Aux.go_X
   #Aux.go_X := #Aux.MidPos_X; (* Convert → Real *)
   // 含义：将 (#Aux.go_X / 1000.0) 赋给 #Aux.go_X
   #Aux.go_X := (#Aux.go_X / 1000.0);
   // 含义：将 SWAP(#StatusIn.go_Z) 赋给 #Aux.MidPos_Z
   #Aux.MidPos_Z := SWAP(#StatusIn.go_Z);
   // 含义：将 #Aux.MidPos_Z; (* Convert → Real *) 赋给 #Aux.go_Z
   #Aux.go_Z := #Aux.MidPos_Z; (* Convert → Real *)
   // 含义：将 (#Aux.go_Z / 1000.0) 赋给 #Aux.go_Z
   #Aux.go_Z := (#Aux.go_Z / 1000.0);

   // ---------- 网络 6 ----------
   // 标题：将用于自定义状态、请求传出
   // 含义：将 "DB1080_Component".Robot.Bus_IN_Data.UserDefineRobOut 赋给 #AtStatusIn
   #AtStatusIn := "DB1080_Component".Robot.Bus_IN_Data.UserDefineRobOut;

   // ---------- 网络 7 ----------
   // 标题：本工位必须要做(可能条件暂时不满足)
   // 含义：当 (#Ctrl_Out.RobotAction = 0) 为 TRUE 时置位 #ChangeTool.OKToStart，否则复位（触点→线圈）
   IF (#Ctrl_Out.RobotAction = 0) THEN
       #ChangeTool.OKToStart := TRUE;
   ELSE
       #ChangeTool.OKToStart := FALSE;
   END_IF;
   // 含义：条件 "ManMode_M" AND "DB1900_Communication_PC".Recv.ChangeToolTPPB 成立时，将 TRUE 传送到 #ChangeTool.StartCmd
   IF "ManMode_M" AND "DB1900_Communication_PC".Recv.ChangeToolTPPB THEN
       #ChangeTool.StartCmd := TRUE;
   END_IF;
   // 含义：条件 NOT (#ChangeTool.StepStart) 成立时，将 0 传送到 "DB1080_Component".Robot.CTRL_IN.ProgNo
   IF NOT (#ChangeTool.StepStart) THEN
       "DB1080_Component".Robot.CTRL_IN.ProgNo := 0;
   END_IF;

   // ---------- 网络 8 ----------
   // 标题：*******************************换夹爪Start****************************************
   // 含义：将 ((((((((((#ChangeTool.StartCmd AND #ChangeTool.OKToStart) OR #ChangeTool.StepStart) AND "AllMode_M") AND "DB1900_Communication_PC".Recv.Z05RetTPPB) AND ("DB1900_Communication_PC".Recv.Current_2 < 0.5))) AND NOT ("DB1040_HomePos".Status.Running)) AND NOT (#ChangeTool.StepEnd)) AND NOT (#ChangeTool.ErrEnd)) AND NOT ("DB1146_PromptFree".ST01.Z07Exting)) AND NOT ("DB1148_PromptBeeper".Public.EMING) 赋给 #ChangeTool.StepStart
   #ChangeTool.StepStart := ((((((((((#ChangeTool.StartCmd AND #ChangeTool.OKToStart) OR #ChangeTool.StepStart) AND "AllMode_M") AND "DB1900_Communication_PC".Recv.Z05RetTPPB) AND ("DB1900_Communication_PC".Recv.Current_2 < 0.5))) AND NOT ("DB1040_HomePos".Status.Running)) AND NOT (#ChangeTool.StepEnd)) AND NOT (#ChangeTool.ErrEnd)) AND NOT ("DB1146_PromptFree".ST01.Z07Exting)) AND NOT ("DB1148_PromptBeeper".Public.EMING);
   // 含义：将 ((((((((((#ChangeTool.StartCmd AND #ChangeTool.OKToStart) OR #ChangeTool.StepStart) AND "AllMode_M") AND "DB1900_Communication_PC".Recv.Z05RetTPPB) AND ("DB1900_Communication_PC".Recv.Current_2 < 0.5))) AND NOT ("DB1040_HomePos".Status.Running)) AND NOT (#ChangeTool.StepEnd)) AND NOT (#ChangeTool.ErrEnd)) AND NOT ("DB1146_PromptFree".ST01.Z07Exting)) AND NOT ("DB1148_PromptBeeper".Public.EMING) 赋给 #ChangeTool.Busy
   #ChangeTool.Busy := ((((((((((#ChangeTool.StartCmd AND #ChangeTool.OKToStart) OR #ChangeTool.StepStart) AND "AllMode_M") AND "DB1900_Communication_PC".Recv.Z05RetTPPB) AND ("DB1900_Communication_PC".Recv.Current_2 < 0.5))) AND NOT ("DB1040_HomePos".Status.Running)) AND NOT (#ChangeTool.StepEnd)) AND NOT (#ChangeTool.ErrEnd)) AND NOT ("DB1146_PromptFree".ST01.Z07Exting)) AND NOT ("DB1148_PromptBeeper".Public.EMING);
   // 含义：将 ((((((((((#ChangeTool.StartCmd AND #ChangeTool.OKToStart) OR #ChangeTool.StepStart) AND "AllMode_M") AND "DB1900_Communication_PC".Recv.Z05RetTPPB) AND ("DB1900_Communication_PC".Recv.Current_2 < 0.5))) AND NOT ("DB1040_HomePos".Status.Running)) AND NOT (#ChangeTool.StepEnd)) AND NOT (#ChangeTool.ErrEnd)) AND NOT ("DB1146_PromptFree".ST01.Z07Exting)) AND NOT ("DB1148_PromptBeeper".Public.EMING) 赋给 "DB1900_Communication_PC".Send.RobotTool
   "DB1900_Communication_PC".Send.RobotTool := ((((((((((#ChangeTool.StartCmd AND #ChangeTool.OKToStart) OR #ChangeTool.StepStart) AND "AllMode_M") AND "DB1900_Communication_PC".Recv.Z05RetTPPB) AND ("DB1900_Communication_PC".Recv.Current_2 < 0.5))) AND NOT ("DB1040_HomePos".Status.Running)) AND NOT (#ChangeTool.StepEnd)) AND NOT (#ChangeTool.ErrEnd)) AND NOT ("DB1146_PromptFree".ST01.Z07Exting)) AND NOT ("DB1148_PromptBeeper".Public.EMING);
   // 含义：条件 NOT (((((((((((#ChangeTool.StartCmd AND #ChangeTool.OKToStart) OR #ChangeTool.StepStart) AND "AllMode_M") AND "DB1900_Communication_PC".Recv.Z05RetTPPB) AND ("DB1900_Communication_PC".Recv.Current_2 < 0.5))) AND NOT ("DB1040_HomePos".Status.Running)) AND NOT (#ChangeTool.StepEnd)) AND NOT (#ChangeTool.ErrEnd)) AND NOT ("DB1146_PromptFree".ST01.Z07Exting)) AND NOT ("DB1148_PromptBeeper".Public.EMING)) 成立时，将 FALSE 传送到 #ChangeTool.ErrEnd
   IF NOT (((((((((((#ChangeTool.StartCmd AND #ChangeTool.OKToStart) OR #ChangeTool.StepStart) AND "AllMode_M") AND "DB1900_Communication_PC".Recv.Z05RetTPPB) AND ("DB1900_Communication_PC".Recv.Current_2 < 0.5))) AND NOT ("DB1040_HomePos".Status.Running)) AND NOT (#ChangeTool.StepEnd)) AND NOT (#ChangeTool.ErrEnd)) AND NOT ("DB1146_PromptFree".ST01.Z07Exting)) AND NOT ("DB1148_PromptBeeper".Public.EMING)) THEN
       #ChangeTool.ErrEnd := FALSE;
   END_IF;

   // ---------- 网络 9 ----------
   // 标题：初始化
   // 含义：条件 (#ChangeTool.StepStart AND NOT (#ChangeTool.ErrEnd)) AND NOT (#ChangeTool.S1) 成立时，将 FALSE 传送到 #ChangeTool.TaskIO
   IF (#ChangeTool.StepStart AND NOT (#ChangeTool.ErrEnd)) AND NOT (#ChangeTool.S1) THEN
       #ChangeTool.TaskIO := FALSE;
   END_IF;
   // 含义：条件 (#ChangeTool.StepStart AND NOT (#ChangeTool.ErrEnd)) AND NOT (#ChangeTool.S1) 成立时，将 FALSE 传送到 #ChangeTool.TaskNIO
   IF (#ChangeTool.StepStart AND NOT (#ChangeTool.ErrEnd)) AND NOT (#ChangeTool.S1) THEN
       #ChangeTool.TaskNIO := FALSE;
   END_IF;
   // 含义：将 #ChangeTool.StepStart AND NOT (#ChangeTool.ErrEnd) 赋给 #ChangeTool.S1
   #ChangeTool.S1 := #ChangeTool.StepStart AND NOT (#ChangeTool.ErrEnd);

   // ---------- 网络 10 ----------
   // 标题：判断条件
   // 含义：条件 #ChangeTool.S1 AND NOT (#ChangeTool.S2) 成立时，将 TRUE 传送到 "DB1081_ValveCall".ST01.Z01.ExtAuto
   IF #ChangeTool.S1 AND NOT (#ChangeTool.S2) THEN
       "DB1081_ValveCall".ST01.Z01.ExtAuto := TRUE;
   END_IF;
   // 含义：条件 #ChangeTool.S1 AND NOT (#ChangeTool.S2) 成立时，将 TRUE 传送到 "DB1081_ValveCall".ST01.Z02.VentValveAuto
   IF #ChangeTool.S1 AND NOT (#ChangeTool.S2) THEN
       "DB1081_ValveCall".ST01.Z02.VentValveAuto := TRUE;
   END_IF;
   // 含义：条件 #ChangeTool.S1 AND NOT (#ChangeTool.S2) 成立时，将 TRUE 传送到 "DB1081_ValveCall".ST01.Z08.ExtAuto
   IF #ChangeTool.S1 AND NOT (#ChangeTool.S2) THEN
       "DB1081_ValveCall".ST01.Z08.ExtAuto := TRUE;
   END_IF;
   // 含义：条件 #ChangeTool.S1 AND NOT (#ChangeTool.S2) 成立时，将 0.4 传送到 "DB1080_Component".Aux.Pressure
   IF #ChangeTool.S1 AND NOT (#ChangeTool.S2) THEN
       "DB1080_Component".Aux.Pressure := 0.4;
   END_IF;
   // 含义：将 ((((#ChangeTool.S1 AND "DB1081_ValveCall".ST01.Z01.ExtPos) AND ("DB1080_Component".ClinyderPos.Ctrl_Out.Cur_Val_Out <= 1.0))) AND "DB1900_Communication_PC".Recv.ParaWriteDone) OR (#ChangeTool.S1 AND #ChangeTool.S2) 赋给 #ChangeTool.S2
   #ChangeTool.S2 := ((((#ChangeTool.S1 AND "DB1081_ValveCall".ST01.Z01.ExtPos) AND ("DB1080_Component".ClinyderPos.Ctrl_Out.Cur_Val_Out <= 1.0))) AND "DB1900_Communication_PC".Recv.ParaWriteDone) OR (#ChangeTool.S1 AND #ChangeTool.S2);

   // ---------- 网络 11 ----------
   // 含义：将 #ChangeTool.S2 AND #ChangeTool.S4 赋给 #ChangeTool.S5
   #ChangeTool.S5 := #ChangeTool.S2 AND #ChangeTool.S4;
   // 含义：将 #ChangeTool.S2 AND #ChangeTool.S3 赋给 #ChangeTool.S4
   #ChangeTool.S4 := #ChangeTool.S2 AND #ChangeTool.S3;
   // 含义：当 #ChangeTool.S2 为 TRUE 时置位 #ChangeTool.S3，否则复位（触点→线圈）
   IF #ChangeTool.S2 THEN
       #ChangeTool.S3 := TRUE;
   ELSE
       #ChangeTool.S3 := FALSE;
   END_IF;

   // ---------- 网络 12 ----------
   // 标题：推力气缸
   // 注释：Thrust Cylinder in Extend Position When Changing Tools, Programmed  By WXY 20230307,
   // 含义：条件 #ChangeTool.S5 AND NOT (#ChangeTool.S7) 成立时，将 TRUE 传送到 "DB1081_ValveCall".ST01.Z05.RetAuto
   IF #ChangeTool.S5 AND NOT (#ChangeTool.S7) THEN
       "DB1081_ValveCall".ST01.Z05.RetAuto := TRUE;
   END_IF;
   // 含义：将 (((((#ChangeTool.S5 AND "IZ02ExtPos") AND "DB1081_ValveCall".ST01.Z01.ExtPos) AND "DB1081_ValveCall".ST01.Z05.RetPos) AND ("DB1080_Component".ClinyderPos.Ctrl_Out.Cur_Val_Out <= 1.0))) OR (#ChangeTool.S5 AND #ChangeTool.S7) 赋给 #ChangeTool.S7
   #ChangeTool.S7 := (((((#ChangeTool.S5 AND "IZ02ExtPos") AND "DB1081_ValveCall".ST01.Z01.ExtPos) AND "DB1081_ValveCall".ST01.Z05.RetPos) AND ("DB1080_Component".ClinyderPos.Ctrl_Out.Cur_Val_Out <= 1.0))) OR (#ChangeTool.S5 AND #ChangeTool.S7);

   // ---------- 网络 13 ----------
   // 含义：将 (#ChangeTool.S7 AND NOT ("DB1080_Component".Robot.Status.Busy)) OR (#ChangeTool.S7 AND #ChangeTool.S10) 赋给 #ChangeTool.S10
   #ChangeTool.S10 := (#ChangeTool.S7 AND NOT ("DB1080_Component".Robot.Status.Busy)) OR (#ChangeTool.S7 AND #ChangeTool.S10);

   // ---------- 网络 14 ----------
   // 标题：快换盘锁紧 253取 254放 左1右2
   // 含义：条件 (#ChangeTool.S10 AND NOT (#ChangeTool.S12)) AND #Aux.ToolAtPosTimer.Q 成立时，将 TRUE 传送到 "DB1080_Component".Robot.Cmd.Auto.ProgStart
   IF (#ChangeTool.S10 AND NOT (#ChangeTool.S12)) AND #Aux.ToolAtPosTimer.Q THEN
       "DB1080_Component".Robot.Cmd.Auto.ProgStart := TRUE;
   END_IF;
   // 含义：条件 (#ChangeTool.S10 AND NOT (#ChangeTool.S12)) AND #Aux.ToolAtPosTimer.Q 成立时，将 254 传送到 "DB1080_Component".Robot.CTRL_IN.ProgNo
   IF (#ChangeTool.S10 AND NOT (#ChangeTool.S12)) AND #Aux.ToolAtPosTimer.Q THEN
       "DB1080_Component".Robot.CTRL_IN.ProgNo := 254;
   END_IF;
   // 含义：条件 ((((#ChangeTool.S10 AND NOT (#ChangeTool.S12)) AND #Aux.ToolAtPosTimer.Q) AND NOT (#Aux.AStation_ToolAtPos)) AND ("DB1080_Component".IOFixtureIID.TP_CurFixtureID = 1)) 成立时，将 1 传送到 #CmdOut.gi_ToolPosNo
   IF ((((#ChangeTool.S10 AND NOT (#ChangeTool.S12)) AND #Aux.ToolAtPosTimer.Q) AND NOT (#Aux.AStation_ToolAtPos)) AND ("DB1080_Component".IOFixtureIID.TP_CurFixtureID = 1)) THEN
       #CmdOut.gi_ToolPosNo := 1;
   END_IF;
   // 含义：条件 ((((#ChangeTool.S10 AND NOT (#ChangeTool.S12)) AND #Aux.ToolAtPosTimer.Q) AND NOT (#Aux.BStation_oolAtPos)) AND ("DB1080_Component".IOFixtureIID.TP_CurFixtureID = 2)) 成立时，将 2 传送到 #CmdOut.gi_ToolPosNo
   IF ((((#ChangeTool.S10 AND NOT (#ChangeTool.S12)) AND #Aux.ToolAtPosTimer.Q) AND NOT (#Aux.BStation_oolAtPos)) AND ("DB1080_Component".IOFixtureIID.TP_CurFixtureID = 2)) THEN
       #CmdOut.gi_ToolPosNo := 2;
   END_IF;
   // 含义：将 (((#ChangeTool.S10 AND NOT (#ChangeTool.S12)) AND #Aux.ToolAtPosTimer.Q) AND #Aux.AStation_ToolAtPosT.Q) AND #Aux.BStation_ToolAtPosT.Q 赋给 "DB1148_PromptBeeper".Public.PutGunPosFull
   "DB1148_PromptBeeper".Public.PutGunPosFull := (((#ChangeTool.S10 AND NOT (#ChangeTool.S12)) AND #Aux.ToolAtPosTimer.Q) AND #Aux.AStation_ToolAtPosT.Q) AND #Aux.BStation_ToolAtPosT.Q;
   // 含义：条件 (#ChangeTool.S10 AND NOT (#ChangeTool.S12)) AND #Aux.ToolAtPosTimer.Q 成立时，将 #CmdOut.gi_ToolPosNo 传送到 #Aux.LastToolPosNo
   IF (#ChangeTool.S10 AND NOT (#ChangeTool.S12)) AND #Aux.ToolAtPosTimer.Q THEN
       #Aux.LastToolPosNo := #CmdOut.gi_ToolPosNo;
   END_IF;
   // 含义：条件 (#ChangeTool.S10 AND NOT (#ChangeTool.S12)) AND #Aux.ToolNotAtPosTimer.Q 成立时，将 TRUE 传送到 "DB1080_Component".Robot.Cmd.Auto.ProgStart
   IF (#ChangeTool.S10 AND NOT (#ChangeTool.S12)) AND #Aux.ToolNotAtPosTimer.Q THEN
       "DB1080_Component".Robot.Cmd.Auto.ProgStart := TRUE;
   END_IF;
   // 含义：条件 (#ChangeTool.S10 AND NOT (#ChangeTool.S12)) AND #Aux.ToolNotAtPosTimer.Q 成立时，将 TRUE 传送到 "DB1081_ValveCall".ST01.Z07.RetAuto
   IF (#ChangeTool.S10 AND NOT (#ChangeTool.S12)) AND #Aux.ToolNotAtPosTimer.Q THEN
       "DB1081_ValveCall".ST01.Z07.RetAuto := TRUE;
   END_IF;
   // 含义：条件 (#ChangeTool.S10 AND NOT (#ChangeTool.S12)) AND #Aux.ToolNotAtPosTimer.Q 成立时，将 253 传送到 "DB1080_Component".Robot.CTRL_IN.ProgNo
   IF (#ChangeTool.S10 AND NOT (#ChangeTool.S12)) AND #Aux.ToolNotAtPosTimer.Q THEN
       "DB1080_Component".Robot.CTRL_IN.ProgNo := 253;
   END_IF;
   // 含义：条件 ((((#ChangeTool.S10 AND NOT (#ChangeTool.S12)) AND #Aux.ToolNotAtPosTimer.Q) AND #Aux.AStation_ToolAtPosT.Q) AND ("DB1900_Communication_PC".Para.IOFixtureNo = 1)) 成立时，将 1 传送到 #CmdOut.gi_ToolPosNo
   IF ((((#ChangeTool.S10 AND NOT (#ChangeTool.S12)) AND #Aux.ToolNotAtPosTimer.Q) AND #Aux.AStation_ToolAtPosT.Q) AND ("DB1900_Communication_PC".Para.IOFixtureNo = 1)) THEN
       #CmdOut.gi_ToolPosNo := 1;
   END_IF;
   // 含义：条件 ((((#ChangeTool.S10 AND NOT (#ChangeTool.S12)) AND #Aux.ToolNotAtPosTimer.Q) AND #Aux.BStation_ToolAtPosT.Q) AND ("DB1900_Communication_PC".Para.IOFixtureNo = 2)) 成立时，将 2 传送到 #CmdOut.gi_ToolPosNo
   IF ((((#ChangeTool.S10 AND NOT (#ChangeTool.S12)) AND #Aux.ToolNotAtPosTimer.Q) AND #Aux.BStation_ToolAtPosT.Q) AND ("DB1900_Communication_PC".Para.IOFixtureNo = 2)) THEN
       #CmdOut.gi_ToolPosNo := 2;
   END_IF;
   // 含义：条件 (((#ChangeTool.S10 AND NOT (#ChangeTool.S12)) AND #Aux.ToolNotAtPosTimer.Q) AND ("DB1900_Communication_PC".Para.IOFixtureNo <> #CmdOut.gi_ToolPosNo)) 成立时，将 TRUE 传送到 "DB1080_Component".Robot.Cmd.Auto.ProgStart
   IF (((#ChangeTool.S10 AND NOT (#ChangeTool.S12)) AND #Aux.ToolNotAtPosTimer.Q) AND ("DB1900_Communication_PC".Para.IOFixtureNo <> #CmdOut.gi_ToolPosNo)) THEN
       "DB1080_Component".Robot.Cmd.Auto.ProgStart := TRUE;
   END_IF;
   // 含义：条件 (((#ChangeTool.S10 AND NOT (#ChangeTool.S12)) AND #Aux.ToolNotAtPosTimer.Q) AND ("DB1900_Communication_PC".Para.IOFixtureNo <> #CmdOut.gi_ToolPosNo)) 成立时，将 TRUE 传送到 #ChangeTool.ErrEnd
   IF (((#ChangeTool.S10 AND NOT (#ChangeTool.S12)) AND #Aux.ToolNotAtPosTimer.Q) AND ("DB1900_Communication_PC".Para.IOFixtureNo <> #CmdOut.gi_ToolPosNo)) THEN
       #ChangeTool.ErrEnd := TRUE;
   END_IF;
   // 含义：将 (((#ChangeTool.S10 AND NOT (#ChangeTool.S12)) AND #Aux.ToolNotAtPosTimer.Q) AND ("DB1900_Communication_PC".Para.IOFixtureNo <> #CmdOut.gi_ToolPosNo)) 赋给 "DB1148_PromptBeeper".Public.FixtureAtPosErr
   "DB1148_PromptBeeper".Public.FixtureAtPosErr := (((#ChangeTool.S10 AND NOT (#ChangeTool.S12)) AND #Aux.ToolNotAtPosTimer.Q) AND ("DB1900_Communication_PC".Para.IOFixtureNo <> #CmdOut.gi_ToolPosNo));
   // 含义：条件 (((((#ChangeTool.S10 AND NOT (#ChangeTool.S12)) AND #Aux.ToolNotAtPosTimer.Q) AND "ManMode_M") AND (#Aux.LastToolPosNo <= 1))) AND #Aux.BStation_ToolAtPosT.Q 成立时，将 2 传送到 #CmdOut.gi_ToolPosNo
   IF (((((#ChangeTool.S10 AND NOT (#ChangeTool.S12)) AND #Aux.ToolNotAtPosTimer.Q) AND "ManMode_M") AND (#Aux.LastToolPosNo <= 1))) AND #Aux.BStation_ToolAtPosT.Q THEN
       #CmdOut.gi_ToolPosNo := 2;
   END_IF;
   // 含义：条件 ((((((#ChangeTool.S10 AND NOT (#ChangeTool.S12)) AND #Aux.ToolNotAtPosTimer.Q) AND "ManMode_M") AND (#Aux.LastToolPosNo <= 1))) AND #Aux.AStation_ToolAtPosT.Q) AND NOT (#Aux.BStation_ToolAtPosT.Q) 成立时，将 1 传送到 #CmdOut.gi_ToolPosNo
   IF ((((((#ChangeTool.S10 AND NOT (#ChangeTool.S12)) AND #Aux.ToolNotAtPosTimer.Q) AND "ManMode_M") AND (#Aux.LastToolPosNo <= 1))) AND #Aux.AStation_ToolAtPosT.Q) AND NOT (#Aux.BStation_ToolAtPosT.Q) THEN
       #CmdOut.gi_ToolPosNo := 1;
   END_IF;
   // 含义：条件 (((((#ChangeTool.S10 AND NOT (#ChangeTool.S12)) AND #Aux.ToolNotAtPosTimer.Q) AND "ManMode_M") AND (#Aux.LastToolPosNo = 2))) AND #Aux.AStation_ToolAtPosT.Q 成立时，将 1 传送到 #CmdOut.gi_ToolPosNo
   IF (((((#ChangeTool.S10 AND NOT (#ChangeTool.S12)) AND #Aux.ToolNotAtPosTimer.Q) AND "ManMode_M") AND (#Aux.LastToolPosNo = 2))) AND #Aux.AStation_ToolAtPosT.Q THEN
       #CmdOut.gi_ToolPosNo := 1;
   END_IF;
   // 含义：条件 ((((((#ChangeTool.S10 AND NOT (#ChangeTool.S12)) AND #Aux.ToolNotAtPosTimer.Q) AND "ManMode_M") AND (#Aux.LastToolPosNo = 2))) AND NOT (#Aux.AStation_ToolAtPosT.Q)) AND #Aux.BStation_ToolAtPosT.Q 成立时，将 2 传送到 #CmdOut.gi_ToolPosNo
   IF ((((((#ChangeTool.S10 AND NOT (#ChangeTool.S12)) AND #Aux.ToolNotAtPosTimer.Q) AND "ManMode_M") AND (#Aux.LastToolPosNo = 2))) AND NOT (#Aux.AStation_ToolAtPosT.Q)) AND #Aux.BStation_ToolAtPosT.Q THEN
       #CmdOut.gi_ToolPosNo := 2;
   END_IF;
   // 含义：条件 #ChangeTool.S10 AND NOT (#ChangeTool.S12) 成立时，将 30 传送到 "DB1080_Component".Robot.CTRL_IN.RobotSpeed
   IF #ChangeTool.S10 AND NOT (#ChangeTool.S12) THEN
       "DB1080_Component".Robot.CTRL_IN.RobotSpeed := 30;
   END_IF;
   // 含义：将 (((((#ChangeTool.S10 AND ("DB1080_Component".Robot.CTRL_IN.ProgNo = 254))) AND NOT (#Aux.AStation_ToolAtPosT.Q)) OR (((#ChangeTool.S10 AND ("DB1080_Component".Robot.CTRL_IN.ProgNo = 254))) AND NOT (#Aux.BStation_ToolAtPosT.Q)) OR (((#ChangeTool.S10 AND ("DB1080_Component".Robot.CTRL_IN.ProgNo = 253))) AND "DB1081_ValveCall".ST01.Z07.RetPos)) AND NOT ("DB1148_PromptBeeper".Public.PutGunPosFull)) OR (#ChangeTool.S10 AND #ChangeTool.S12) 赋给 #ChangeTool.S12
   #ChangeTool.S12 := (((((#ChangeTool.S10 AND ("DB1080_Component".Robot.CTRL_IN.ProgNo = 254))) AND NOT (#Aux.AStation_ToolAtPosT.Q)) OR (((#ChangeTool.S10 AND ("DB1080_Component".Robot.CTRL_IN.ProgNo = 254))) AND NOT (#Aux.BStation_ToolAtPosT.Q)) OR (((#ChangeTool.S10 AND ("DB1080_Component".Robot.CTRL_IN.ProgNo = 253))) AND "DB1081_ValveCall".ST01.Z07.RetPos)) AND NOT ("DB1148_PromptBeeper".Public.PutGunPosFull)) OR (#ChangeTool.S10 AND #ChangeTool.S12);

   // ---------- 网络 15 ----------
   // 标题：右防尘盖夹紧缸
   // 含义：条件 ((#ChangeTool.S12 AND NOT (#ChangeTool.S13)) AND (#CmdOut.gi_ToolPosNo = 1)) 成立时，将 TRUE 传送到 "DB1081_ValveCall".ST01.Z03.ExtAuto
   IF ((#ChangeTool.S12 AND NOT (#ChangeTool.S13)) AND (#CmdOut.gi_ToolPosNo = 1)) THEN
       "DB1081_ValveCall".ST01.Z03.ExtAuto := TRUE;
   END_IF;
   // 含义：条件 ((#ChangeTool.S12 AND NOT (#ChangeTool.S13)) AND (#CmdOut.gi_ToolPosNo = 2)) 成立时，将 TRUE 传送到 "DB1081_ValveCall".ST01.Z04.ExtAuto
   IF ((#ChangeTool.S12 AND NOT (#ChangeTool.S13)) AND (#CmdOut.gi_ToolPosNo = 2)) THEN
       "DB1081_ValveCall".ST01.Z04.ExtAuto := TRUE;
   END_IF;
   // 含义：条件 (((((#ChangeTool.S12 AND NOT (#ChangeTool.S13)) AND ("DB1080_Component".Robot.CTRL_IN.ProgNo = 254))) OR (((#ChangeTool.S12 AND NOT (#ChangeTool.S13)) AND ("DB1080_Component".Robot.CTRL_IN.ProgNo = 253)))) AND (#CmdOut.gi_ToolPosNo = 1)) 成立时，将 TRUE 传送到 "DB1081_ValveCall".ST01.Z03.ExtAuto
   IF (((((#ChangeTool.S12 AND NOT (#ChangeTool.S13)) AND ("DB1080_Component".Robot.CTRL_IN.ProgNo = 254))) OR (((#ChangeTool.S12 AND NOT (#ChangeTool.S13)) AND ("DB1080_Component".Robot.CTRL_IN.ProgNo = 253)))) AND (#CmdOut.gi_ToolPosNo = 1)) THEN
       "DB1081_ValveCall".ST01.Z03.ExtAuto := TRUE;
   END_IF;
   // 含义：条件 (((((#ChangeTool.S12 AND NOT (#ChangeTool.S13)) AND ("DB1080_Component".Robot.CTRL_IN.ProgNo = 254))) OR (((#ChangeTool.S12 AND NOT (#ChangeTool.S13)) AND ("DB1080_Component".Robot.CTRL_IN.ProgNo = 253)))) AND (#CmdOut.gi_ToolPosNo = 2)) 成立时，将 TRUE 传送到 "DB1081_ValveCall".ST01.Z04.ExtAuto
   IF (((((#ChangeTool.S12 AND NOT (#ChangeTool.S13)) AND ("DB1080_Component".Robot.CTRL_IN.ProgNo = 254))) OR (((#ChangeTool.S12 AND NOT (#ChangeTool.S13)) AND ("DB1080_Component".Robot.CTRL_IN.ProgNo = 253)))) AND (#CmdOut.gi_ToolPosNo = 2)) THEN
       "DB1081_ValveCall".ST01.Z04.ExtAuto := TRUE;
   END_IF;
   // 含义：将 (((((((((#ChangeTool.S12 AND ("DB1080_Component".Robot.CTRL_IN.ProgNo = 254))) AND (#CmdOut.gi_ToolPosNo = 1))) AND NOT (#Aux.AStation_ToolAtPosT.Q)) OR (((((#ChangeTool.S12 AND ("DB1080_Component".Robot.CTRL_IN.ProgNo = 254))) AND (#CmdOut.gi_ToolPosNo = 2))) AND NOT (#Aux.BStation_ToolAtPosT.Q)) OR ((#ChangeTool.S12 AND ("DB1080_Component".Robot.CTRL_IN.ProgNo = 253)))) AND (#CmdOut.gi_ToolPosNo = 2))) AND "DB1081_ValveCall".ST01.Z04.ExtPos) OR (((((((((#ChangeTool.S12 AND ("DB1080_Component".Robot.CTRL_IN.ProgNo = 254))) AND (#CmdOut.gi_ToolPosNo = 1))) AND NOT (#Aux.AStation_ToolAtPosT.Q)) OR (((((#ChangeTool.S12 AND ("DB1080_Component".Robot.CTRL_IN.ProgNo = 254))) AND (#CmdOut.gi_ToolPosNo = 2))) AND NOT (#Aux.BStation_ToolAtPosT.Q)) OR ((#ChangeTool.S12 AND ("DB1080_Component".Robot.CTRL_IN.ProgNo = 253)))) AND (#CmdOut.gi_ToolPosNo = 1))) AND "DB1081_ValveCall".ST01.Z03.ExtPos) OR (#ChangeTool.S12 AND #ChangeTool.S13) 赋给 #ChangeTool.S13
   #ChangeTool.S13 := (((((((((#ChangeTool.S12 AND ("DB1080_Component".Robot.CTRL_IN.ProgNo = 254))) AND (#CmdOut.gi_ToolPosNo = 1))) AND NOT (#Aux.AStation_ToolAtPosT.Q)) OR (((((#ChangeTool.S12 AND ("DB1080_Component".Robot.CTRL_IN.ProgNo = 254))) AND (#CmdOut.gi_ToolPosNo = 2))) AND NOT (#Aux.BStation_ToolAtPosT.Q)) OR ((#ChangeTool.S12 AND ("DB1080_Component".Robot.CTRL_IN.ProgNo = 253)))) AND (#CmdOut.gi_ToolPosNo = 2))) AND "DB1081_ValveCall".ST01.Z04.ExtPos) OR (((((((((#ChangeTool.S12 AND ("DB1080_Component".Robot.CTRL_IN.ProgNo = 254))) AND (#CmdOut.gi_ToolPosNo = 1))) AND NOT (#Aux.AStation_ToolAtPosT.Q)) OR (((((#ChangeTool.S12 AND ("DB1080_Component".Robot.CTRL_IN.ProgNo = 254))) AND (#CmdOut.gi_ToolPosNo = 2))) AND NOT (#Aux.BStation_ToolAtPosT.Q)) OR ((#ChangeTool.S12 AND ("DB1080_Component".Robot.CTRL_IN.ProgNo = 253)))) AND (#CmdOut.gi_ToolPosNo = 1))) AND "DB1081_ValveCall".ST01.Z03.ExtPos) OR (#ChangeTool.S12 AND #ChangeTool.S13);

   // ---------- 网络 16 ----------
   // 标题：调用机器人
   // 含义：条件 #ChangeTool.S13 AND NOT (#ChangeTool.S15) 成立时，将 TRUE 传送到 "DB1080_Component".Robot.Cmd.Auto.ProgStart
   IF #ChangeTool.S13 AND NOT (#ChangeTool.S15) THEN
       "DB1080_Component".Robot.Cmd.Auto.ProgStart := TRUE;
   END_IF;
   // 含义：将 #ChangeTool.S13 AND NOT (#ChangeTool.S15) 赋给 "DB1146_PromptFree".Public.do_ChgGrp_Act
   "DB1146_PromptFree".Public.do_ChgGrp_Act := #ChangeTool.S13 AND NOT (#ChangeTool.S15);
   // 含义：将 ((#ChangeTool.S13 AND "DB1080_Component".Robot.Status.Busy) AND #StatusIn.do_ChgGrp_Act) OR (#ChangeTool.S13 AND #ChangeTool.S15) 赋给 #ChangeTool.S15
   #ChangeTool.S15 := ((#ChangeTool.S13 AND "DB1080_Component".Robot.Status.Busy) AND #StatusIn.do_ChgGrp_Act) OR (#ChangeTool.S13 AND #ChangeTool.S15);

